(* IEC 61131-3 sources: stdmachine/plc/src/05_Sequencers (part 2) *)

(* ---- FB_Machine.st ---- *)
// Bloc de tête du PLC (docs/05 § 5.1, § 5.2, § 10 ; docs/06 § 6) : machine d'états de la machine, propagation des
// commandes aux stations, défauts machine et raison d'arrêt, objets de niveau machine, système planaire, séquenceur
// général, calibrations machine, chargeur, handshakes de GVL_Hmi, forçages, surveillance des rebuts, balise,
// identité du PLC, battement de la HMI, publication du statut.
//
// Le projet de la machine l'appelle une fois par cycle dans MAIN : fbMachine(); après avoir renseigné GVL_IoRef.
// Avant le premier appel, il peut donner ses pools (SetPools) et son pilote planaire (SetPlanarDriver) ; sinon la
// bibliothèque prend FB_DefaultPools et le système planaire simulé.
FUNCTION_BLOCK FB_Machine EXTENDS FB_NodeBase IMPLEMENTS I_ManualHost, I_ObjectHost
VAR
    fbPack : FB_PackML;
    aStation : ARRAY[1..GVL_Const.MAX_STATIONS] OF FB_Station;
    fbSeq : FB_GeneralSequencer;
    fbMgr : FB_MoverManager;
    fbPlanarSim : FB_PlanarSim;
    fbAlarms : FB_AlarmManager;
    fbTraces : FB_TraceBuffer;
    fbQuality : FB_QualityMonitor;
    fbFactory : FB_ObjectFactory;
    fbLoader : FB_Loader;
    fbCalib : FB_MachineCalib;
    fbDefaultPools : FB_DefaultPools;
    fbManual : FB_ManualChannel;            // canal 0 : objets de niveau machine
    _ipPools : I_ObjectPools;
    _ipPlanar : I_PlanarDriver;
    _bSimPlanar : BOOL;
    aObj : ARRAY[1..GVL_Const.MAX_MACHINE_OBJ] OF I_Object;
    _nObj : UINT;
    _bInit : BOOL;
    _ePendingCmd : E_Cmd;
    _sCmdUser : STRING(24);
    _eReasonNext : E_StopReason;            // cause système du prochain arrêt
    _bOperatorAwaited : BOOL;               // fin d'OF, machine vidée : bleu clignotant jusqu'au prochain Start
    // Handshakes (docs/06 § 6.1) : dernier nSeq traité
    _nCmdSeq : UDINT;
    _nOverrideSeq : UDINT;
    _nLaunchSeq : UDINT;
    _nOrderSeq : UDINT;
    _nMoverVarSeq : UDINT;
    _nPromptSeq : UDINT;
    _nPartSeq : UDINT;
    _nAckSeq : UDINT;
    _nForceSeq : UDINT;
    _nQualitySeq : UDINT;
    _nSimForceSeq : UDINT;
    // Battement de la HMI
    _nLastHmiBeat : UDINT;
    _fHmiQuietMs : LREAL;
    bHmiLost : BOOL;
    _nHeartbeat : UDINT;
    _fRetainedMs : LREAL;
    _tLastCalibCheck : LINT;
    _nPlanarError : UINT;
END_VAR
VAR PERSISTENT
    stForce : ST_MachineForce;              // forçages et état déclaré (docs/12)
    _fMachineOverride : LREAL := 100.0;
    _aStationOverride : ARRAY[1..GVL_Const.MAX_STATIONS] OF LREAL := [16(100.0)];
    _eMode : E_Mode;
    _nStopCauseGid : UDINT;
    _nStopCauseCode : UINT;
    _eStopReason : E_StopReason;
END_VAR

_Run();

// ================================================================== mise en place

METHOD SetPools
VAR_INPUT
    ipPools : I_ObjectPools;
END_VAR
_ipPools := ipPools;
END_METHOD

METHOD SetPlanarDriver
VAR_INPUT
    ipDriver : I_PlanarDriver;
END_VAR
_ipPlanar := ipDriver;
END_METHOD

METHOD PRIVATE _Init
VAR
    n : USINT;
    t : UINT;
    stResp : ST_DeployResponse;
END_VAR
fbAlarms.Bind(GVL_Hmi.stAlarms);
fbTraces.Bind(GVL_Hmi.stTraces);
IF _ipPools = 0 THEN _ipPools := fbDefaultPools; END_IF
IF _ipPlanar = 0 THEN
    _ipPlanar := fbPlanarSim;
    _bSimPlanar := TRUE;
END_IF
fbFactory.SetPools(_ipPools, fbAlarms);
fbFactory.SetHost(0, THIS^, THIS^, 0);
FOR n := 1 TO GVL_Const.MAX_STATIONS DO
    aStation[n].Init(nStation := n, refData := GVL_Active.aStation[n], refMachine := GVL_Active.stMachine, refAlarms := fbAlarms,
                     refStatus := GVL_Hmi.aStationStatus[n], refStep := GVL_Hmi.aStep[n], ipMachine := THIS^);
    aStation[n].SetOverride(_aStationOverride[n]);
    fbFactory.SetHost(n, aStation[n], aStation[n], aStation[n]);
    fbSeq.SetStation(n, ADR(aStation[n]));
    fbCalib.SetStation(n, ADR(aStation[n]));
END_FOR
fbQuality.Init(GVL_Active.stMachine, fbAlarms);
fbMgr.Init(GVL_Active.stMachine, _ipPlanar);
GVL_IoRef.ipPlanar := _ipPlanar;
GVL_IoRef.ipMovers := fbMgr;
fbSeq.Init(GVL_Active.stMachine, fbMgr, fbQuality, fbAlarms, fbTraces);
fbCalib.Init(GVL_Active.stMachine, fbAlarms, fbMgr);
fbManual.Init(nStation := 0, ipHost := THIS^);
fbLoader.Init(fbFactory);
SetOverride(_fMachineOverride);

// Mémoire rémanente : identifiant tiré à sa première initialisation (docs/02 § 7.4)
IF GVL_Active.nRetainId = 0 THEN
    GVL_Active.nRetainId := LINT_TO_ULINT(F_NowUtc()) XOR 16#9E3779B97F4A7C15;
END_IF

// Redémarrage du PLC : le dernier déploiement reste actif, les objets sont rattachés de nouveau à leurs éléments
IF GVL_Active.bDeployed THEN
    fbFactory.Build(stResp);
    fbMgr.Configure();
    fbSeq.ScanGroups();
    _PlaceSimMovers();
END_IF
FOR n := 1 TO GVL_Const.MAX_STATIONS DO aStation[n].SetMode(_eMode); END_FOR

// Identité (docs/05 § 10)
GVL_Hmi.stIdentity.nInterfaceVersion := GVL_Const.INTERFACE_VERSION;
GVL_Hmi.stIdentity.nInstrSetVersion := GVL_Const.INSTR_SET_VERSION;
GVL_Hmi.stIdentity.nCatalogVersion := GVL_Catalog.CatalogVersion;
GVL_Hmi.stIdentity.sLibVersion := GVL_Const.LIB_VERSION;
GVL_Hmi.stIdentity.nRetainId := GVL_Active.nRetainId;
FOR t := 1 TO GVL_Const.MAX_TYPE DO GVL_Hmi.stIdentity.aPoolSize[t] := fbFactory.PoolSize(t); END_FOR

// Les demandes déjà présentes dans GVL_Hmi au démarrage ne sont pas rejouées
_nCmdSeq := GVL_Hmi.stCmd.nSeq;
_nOverrideSeq := GVL_Hmi.stOverride.nSeq;
_nLaunchSeq := GVL_Hmi.stLaunch.nSeq;
_nOrderSeq := GVL_Hmi.stOrder.nSeq;
_nMoverVarSeq := GVL_Hmi.stMoverVar.nSeq;
_nPromptSeq := GVL_Hmi.stPrompt.nSeq;
_nPartSeq := GVL_Hmi.stPartCmd.nSeq;
_nAckSeq := GVL_Hmi.stAlarmAck.nSeq;
_nForceSeq := GVL_Hmi.stForceCmd.nSeq;
_nQualitySeq := GVL_Hmi.stQualityCmd.nSeq;
_nSimForceSeq := GVL_Hmi.stSimForce.nSeq;
_nLastHmiBeat := GVL_Hmi.nHmiHeartbeat;
_ApplyMoverForces();
_bInit := TRUE;
END_METHOD

// Simulation : chaque mover est posé sur une position tampon, sinon de parcage, sinon en ligne (docs/06 § 8)
METHOD PRIVATE _PlaceSimMovers
VAR
    i : USINT;
    k : INT;
    nPlaced : USINT;
    stPos : ST_Position;
END_VAR
IF NOT _bSimPlanar THEN RETURN; END_IF
fbPlanarSim.SetMoverCount(GVL_Active.stMachine.nMovers);
nPlaced := 0;
FOR k := 1 TO GVL_Active.stMachine.nPlanarPos DO
    IF nPlaced < GVL_Active.stMachine.nMovers AND (GVL_Active.stMachine.aPlanarPos[k].eKind = E_PlanarPosKind.Buffer
       OR GVL_Active.stMachine.aPlanarPos[k].eKind = E_PlanarPosKind.Park) THEN
        nPlaced := nPlaced + 1;
        fbPlanarSim.SetInitialPosition(nPlaced, GVL_Active.stMachine.aPlanarPos[k].stPos);
    END_IF
END_FOR
FOR i := nPlaced + 1 TO GVL_Active.stMachine.nMovers DO
    MEMSET(ADR(stPos), 0, SIZEOF(stPos));
    stPos.fX := USINT_TO_LREAL(i) * 120.0;
    fbPlanarSim.SetInitialPosition(i, stPos);
END_FOR
END_METHOD

// ================================================================== cycle

METHOD PRIVATE _Run
VAR
    n : USINT;
    k : UINT;
    eBefore : E_State;
    eCmd : E_Cmd;
    tNow : LINT;
END_VAR
IF NOT _bInit THEN _Init(); END_IF
tNow := F_NowUtc();
_nHeartbeat := _nHeartbeat + 1;
_WatchHmi();

// Chargeur : vérification, activation, restauration (machine Stopped)
fbLoader(bMachineStopped := fbPack.eState = E_State.Stopped);
fbLoader.Cycle();
IF fbLoader.bActivate THEN _Activate(); END_IF
IF fbLoader.bRestore THEN _ApplyRestore(); END_IF

// Demandes de la HMI
_HandleCmd();
_HandleOverride();
_HandleLaunch();
_HandleOrder();
_HandleMoverVar();
_HandlePrompt();
_HandlePart();
_HandleAlarmAck();
_HandleForce();
_HandleQuality();
_HandleSimForce();

// Arrêts automatiques demandés au cycle précédent : OF terminé, machine vidée, réaction qualité
IF fbSeq.bStopRequest AND _ePendingCmd = E_Cmd.None AND fbPack.Accepts(E_Cmd.Stop) THEN
    _ePendingCmd := E_Cmd.Stop;
    CASE fbSeq.nStopReason OF
        1: _eReasonNext := E_StopReason.OrderComplete;
        2: _eReasonNext := E_StopReason.Drained;
    ELSE
        _eReasonNext := E_StopReason.Quality;
    END_CASE
    _bOperatorAwaited := fbSeq.nStopReason <> 3;
END_IF

// Système planaire
UpdateOverride();
fbMgr.Cycle(EffectiveOverride);         // fait aussi tourner le pilote planaire
_PlanarAlarms();

// Machine d'états
eCmd := _ePendingCmd;
_ePendingCmd := E_Cmd.None;
eBefore := fbPack.eState;
fbPack(eCmd := eCmd, bStateComplete := _StateComplete(), bFault := _Fault());
IF fbPack.bEntry THEN _OnEntry(eBefore); END_IF

// Objets de niveau machine
_UpdateObjects();
fbManual.Cycle();

// Stations : forçages et réactions qualité, puis leur cycle
FOR n := 1 TO GVL_Const.MAX_STATIONS DO
    aStation[n].SetOutOfProduction(stForce.aStation[n].bOutOfProduction);
    aStation[n].SetQualityLock(fbQuality.aStationHold[n]);
    aStation[n].Cycle();
END_FOR

// Séquenceur général et calibration machine
fbSeq.Cycle(fbPack.eState);
IF fbCalib.bRunning AND (fbPack.eState <> E_State.Idle OR _eMode <> E_Mode.Maintenance) THEN fbCalib.Abort(); END_IF
fbCalib.Cycle(bHmiLost);

// Calibrations échues : une fois par jour (et à chaque Reset, voir _OnEntry)
IF tNow - _tLastCalibCheck > 864000000000 THEN _CheckCalibrations(tNow); END_IF

_Beacon();
fbQuality.Publish();
_fRetainedMs := _fRetainedMs + F_CycleMs();
IF _fRetainedMs >= 1000.0 THEN
    _fRetainedMs := 0;
    _PublishRetained();
END_IF
_Publish();
END_METHOD

METHOD PRIVATE _WatchHmi
IF GVL_Hmi.nHmiHeartbeat <> _nLastHmiBeat THEN
    _nLastHmiBeat := GVL_Hmi.nHmiHeartbeat;
    _fHmiQuietMs := 0;
    bHmiLost := FALSE;
ELSE
    _fHmiQuietMs := _fHmiQuietMs + F_CycleMs();
    IF _fHmiQuietMs >= GVL_Const.HMI_HEARTBEAT_MS AND NOT bHmiLost THEN
        bHmiLost := TRUE;
        fbAlarms.RaiseEvent(0, 917, 0, E_Severity.Info);           // la production continue (docs/06 § 6.2)
    END_IF
END_IF
END_METHOD

// ================================================================== machine d'états (docs/05 § 5.1 et 5.2)

METHOD PRIVATE _StateComplete : BOOL
VAR
    n : USINT;
    bAll : BOOL := TRUE;
END_VAR
_StateComplete := FALSE;
CASE fbPack.eState OF
    E_State.Resetting:
        // Système planaire actif, movers détectés (un mover hors service peut être absent), chaque fonction
        // utilisée a une station en Idle
        IF NOT _ipPlanar.Activate(TRUE) THEN RETURN; END_IF
        _StateComplete := _AllMoversDetected() AND fbSeq.MissingGroup(2) = 0;
    E_State.Stopping:
        FOR n := 1 TO GVL_Const.MAX_STATIONS DO
            IF aStation[n].State <> E_State.Stopped AND aStation[n].State <> E_State.Aborted THEN bAll := FALSE; END_IF
        END_FOR
        _StateComplete := bAll AND NOT fbMgr.AnyMoving();
    E_State.Clearing:
        FOR n := 1 TO GVL_Const.MAX_STATIONS DO
            IF aStation[n].State = E_State.Clearing THEN bAll := FALSE; END_IF
        END_FOR
        _StateComplete := bAll AND _ObjectsOk();
END_CASE
END_METHOD

METHOD PRIVATE _AllMoversDetected : BOOL
VAR
    i : USINT;
END_VAR
_AllMoversDetected := TRUE;
FOR i := 1 TO GVL_Active.stMachine.nMovers DO
    IF NOT _ipPlanar.MoverDetected(i) THEN
        IF NOT stForce.aMover[i].bOutOfService THEN
            _AllMoversDetected := FALSE;
            fbAlarms.Raise(_PlanarGlobalId(), 101, i, E_Severity.Warning);    // « Mover non détecté » : reste en Resetting
        END_IF
    ELSE
        fbAlarms.Clear(_PlanarGlobalId(), 101);
    END_IF
END_FOR
END_METHOD

METHOD PRIVATE _Fault : BOOL
VAR
    n : USINT;
    g : USINT;
    eSt : E_State;
    ipSafety : I_SafetyCircuits;
    k : UINT;
END_VAR
_Fault := FALSE;
eSt := fbPack.eState;
// Circuits de sécurité de niveau machine
FOR k := 1 TO _nObj DO
    IF aObj[k] <> 0 AND_THEN __QUERYINTERFACE(aObj[k], ipSafety) THEN
        IF NOT ipSafety.AllOk THEN _Fault := TRUE; END_IF
    END_IF
END_FOR
IF eSt = E_State.Stopped THEN RETURN; END_IF          // à l'arrêt, une sécurité ouverte n'est pas un défaut
// Système planaire, movers, alarmes de process de gravité défaut machine
IF _nPlanarError <> 0 OR fbSeq.bMachineFault THEN _Fault := TRUE; END_IF
IF eSt <> E_State.Aborted AND eSt <> E_State.Clearing THEN
    FOR n := 1 TO GVL_Const.MAX_STATIONS DO
        IF aStation[n].MachineFault THEN _Fault := TRUE; END_IF
    END_FOR
    IF NOT _ObjectsOk() THEN _Fault := TRUE; END_IF
END_IF
// Fonction utilisée sans station disponible (913) ; au Reset, fonction dont toutes les stations ont échoué
IF eSt = E_State.Execute THEN
    g := fbSeq.MissingGroup(1);
ELSIF eSt = E_State.Resetting THEN
    g := fbSeq.MissingGroup(3);
END_IF
IF g <> 0 THEN
    fbAlarms.RaiseEvent(0, 913, g, E_Severity.MachineFault);
    _Fault := TRUE;
END_IF
END_METHOD

METHOD PRIVATE _ObjectsOk : BOOL
VAR
    k : UINT;
END_VAR
_ObjectsOk := TRUE;
FOR k := 1 TO _nObj DO
    IF aObj[k] <> 0 THEN
        IF aObj[k].NodeState = E_ObjState.Error THEN _ObjectsOk := FALSE; END_IF
    END_IF
END_FOR
END_METHOD

METHOD PRIVATE _OnEntry
VAR_INPUT
    eFrom : E_State;
END_VAR
VAR
    n : USINT;
    k : UINT;
    eSt : E_State;
END_VAR
CASE fbPack.eState OF
    E_State.Stopped:
        fbSeq.bDrain := FALSE;
    E_State.Resetting:
        _ClearStopCause();
        FOR k := 1 TO _nObj DO IF aObj[k] <> 0 THEN aObj[k].Ack(); END_IF END_FOR
        _ipPlanar.AckError();
        FOR n := 1 TO GVL_Const.MAX_STATIONS DO
            IF _StationUsed(n) AND aStation[n].State = E_State.Stopped THEN aStation[n].Command(E_Cmd.Reset); END_IF
        END_FOR
        _CheckCalibrations(F_NowUtc());
    E_State.Idle:
        // Fin du Reset : chaque mover reçoit sa position, contextes et pièces gardés (docs/05 § 6.3)
        IF eFrom = E_State.Resetting THEN fbSeq.OnReset(); END_IF
    E_State.Execute:
        _ClearStopCause();
        _bOperatorAwaited := FALSE;
        FOR n := 1 TO GVL_Const.MAX_STATIONS DO
            eSt := aStation[n].State;
            IF _StationUsed(n) AND (eSt = E_State.Idle OR eSt = E_State.Held) THEN aStation[n].Command(E_Cmd.Start); END_IF
        END_FOR
    E_State.Held:
        _TakeStopCause();
        FOR n := 1 TO GVL_Const.MAX_STATIONS DO
            IF aStation[n].State = E_State.Execute THEN aStation[n].Command(E_Cmd.Hold); END_IF
        END_FOR
    E_State.Stopping:
        _TakeStopCause();
        fbSeq.bDrain := FALSE;
        FOR n := 1 TO GVL_Const.MAX_STATIONS DO
            eSt := aStation[n].State;
            IF eSt = E_State.Resetting OR eSt = E_State.Idle OR eSt = E_State.Execute OR eSt = E_State.Held THEN aStation[n].Command(E_Cmd.Stop); END_IF
        END_FOR
    E_State.Aborted:
        _TakeStopCause();
        fbSeq.bDrain := FALSE;
        fbMgr.StopAll();
        fbCalib.Abort();
        FOR k := _nObj TO 1 BY -1 DO IF aObj[k] <> 0 THEN aObj[k].Abort(); END_IF END_FOR
        FOR n := 1 TO GVL_Const.MAX_STATIONS DO
            IF aStation[n].State <> E_State.Aborted AND aStation[n].State <> E_State.Stopped THEN aStation[n].Command(E_Cmd.Abort); END_IF
        END_FOR
    E_State.Clearing:
        fbAlarms.AckFaults(0, FALSE, _sCmdUser);
        FOR k := 1 TO _nObj DO IF aObj[k] <> 0 THEN aObj[k].Ack(); END_IF END_FOR
        fbSeq.ClearFaults();
        _ipPlanar.AckError();
        FOR n := 1 TO GVL_Const.MAX_STATIONS DO
            IF aStation[n].State = E_State.Aborted THEN aStation[n].Command(E_Cmd.Clear); END_IF
        END_FOR
END_CASE
END_METHOD

METHOD PRIVATE _StationUsed : BOOL
VAR_INPUT
    n : USINT;
END_VAR
_StationUsed := GVL_Active.stMachine.aStation[n].bUsed;
END_METHOD

// Raison d'arrêt (docs/05 § 5.2, docs/14 § 4) : première alarme cause, sinon la cause système
METHOD PRIVATE _TakeStopCause
VAR
    i : INT;
END_VAR
IF _eStopReason <> E_StopReason.None THEN RETURN; END_IF      // déjà prise pour cet épisode d'arrêt
// Un arrêt automatique (OF terminé, machine vidée, qualité) garde sa cause même si une alarme est active
IF _eReasonNext = E_StopReason.OrderComplete OR _eReasonNext = E_StopReason.Drained OR _eReasonNext = E_StopReason.Quality THEN
    _eStopReason := _eReasonNext;
    _eReasonNext := E_StopReason.None;
    RETURN;
END_IF
i := fbAlarms.FirstFault(0, TRUE);
IF i > 0 THEN
    fbAlarms.MarkCause(i);
    _nStopCauseGid := GVL_Hmi.stAlarms.aActive[i].nGlobalId;
    _nStopCauseCode := GVL_Hmi.stAlarms.aActive[i].nCode;
    _eStopReason := E_StopReason.Alarm;
ELSE
    _eStopReason := E_StopReason.Operator;
END_IF
_eReasonNext := E_StopReason.None;
END_METHOD

METHOD PRIVATE _ClearStopCause
_nStopCauseGid := 0;
_nStopCauseCode := 0;
_eStopReason := E_StopReason.None;
_eReasonNext := E_StopReason.None;
END_METHOD

METHOD PRIVATE _CheckCalibrations
VAR_INPUT
    tNow : LINT;
END_VAR
VAR
    n : USINT;
END_VAR
_tLastCalibCheck := tNow;
FOR n := 1 TO GVL_Const.MAX_STATIONS DO
    IF _StationUsed(n) THEN aStation[n].CheckCalibrations(tNow); END_IF
END_FOR
fbCalib.CheckCalibrations(tNow);
END_METHOD

// ================================================================== système planaire et objets machine

METHOD PRIVATE _PlanarGlobalId : UDINT
VAR
    k : UINT;
END_VAR
_PlanarGlobalId := 0;
FOR k := 1 TO MIN(GVL_Active.stMachine.nMachineObj, GVL_Const.MAX_MACHINE_OBJ) DO
    IF GVL_Active.stMachine.aMachineObj[k].nType = GVL_Catalog.Type_PlanarSystem THEN
        _PlanarGlobalId := UINT_TO_UDINT(GVL_Active.stMachine.aMachineObj[k].nLocalId);
        RETURN;
    END_IF
END_FOR
END_METHOD

METHOD PRIVATE _PlanarAlarms
VAR
    nErr : UINT;
END_VAR
nErr := _ipPlanar.ErrorCode;
IF nErr <> _nPlanarError THEN
    IF _nPlanarError <> 0 THEN fbAlarms.Clear(_PlanarGlobalId(), _nPlanarError); END_IF
    IF nErr <> 0 THEN fbAlarms.Raise(_PlanarGlobalId(), nErr, _ipPlanar.ErrorSubCode, E_Severity.MachineFault); END_IF
    _nPlanarError := nErr;
END_IF
END_METHOD

METHOD PRIVATE _UpdateObjects
VAR
    k : UINT;
END_VAR
FOR k := 1 TO _nObj DO
    IF aObj[k] <> 0 THEN
        aObj[k].Cycle();
        GVL_Hmi.aObjStatus[0, k] := aObj[k].Status;
    END_IF
END_FOR
END_METHOD

// Balise de la machine (docs/02 § 8) : pilotée par l'état de la machine
METHOD PRIVATE _Beacon
VAR
    k : UINT;
    n : USINT;
    nPattern : UINT;
    bMaint : BOOL;
    bStationAborted : BOOL;
    ipBeacon : I_Beacon;
END_VAR
bMaint := _eMode = E_Mode.Maintenance OR stForce.eDeclared = E_DeclaredState.PlannedMaintenance
          OR stForce.eDeclared = E_DeclaredState.CorrectiveMaintenance OR stForce.eDeclared = E_DeclaredState.Trials
          OR stForce.eDeclared = E_DeclaredState.Cleaning;
FOR n := 1 TO GVL_Const.MAX_STATIONS DO
    IF aStation[n].State = E_State.Aborted THEN bStationAborted := TRUE; END_IF
END_FOR
nPattern := F_BeaconPattern(fbPack.eState, bMaint, _bOperatorAwaited OR fbSeq.AnyToEmpty() OR fbQuality.bAnyReaction, bStationAborted);
FOR k := 1 TO _nObj DO
    IF aObj[k] <> 0 AND_THEN __QUERYINTERFACE(aObj[k], ipBeacon) THEN ipBeacon.SetPattern(nPattern, (nPattern AND GVL_BeaconBits.BUZZER) <> 0); END_IF
END_FOR
END_METHOD

// ================================================================== déploiement (docs/05 § 10)

METHOD PRIVATE _Activate
VAR
    stResp : ST_DeployResponse;
    n : USINT;
    nOldGeneral : INT;
    nNewGeneral : INT;
    bRestart : BOOL;
END_VAR
IF fbPack.eState <> E_State.Stopped THEN
    F_AddDeployError(stResp, 21, 0, 0, 0, 0, 0);
    fbLoader.Finish(stResp);
    RETURN;
END_IF
nOldGeneral := _GeneralSize(GVL_Active.stMachine);
nNewGeneral := _GeneralSize(GVL_Hmi.stStaging.stMachine);
bRestart := NOT GVL_Active.bDeployed OR nOldGeneral <> nNewGeneral
            OR GVL_Active.stMachine.nMovers <> GVL_Hmi.stStaging.stMachine.nMovers
            OR GVL_Active.stMachine.nSlots <> GVL_Hmi.stStaging.stMachine.nSlots;
// Copie atomique de la zone d'attente (un seul cycle)
GVL_Active.stMachine := GVL_Hmi.stStaging.stMachine;
GVL_Active.aStation := GVL_Hmi.stStaging.aStation;
GVL_Active.aPressRecipe := GVL_Hmi.stStaging.aPressRecipe;
GVL_Active.stMachine.tDeployed := F_NowUtc();
GVL_Active.stMachine.sDeployedBy := fbLoader.Request.sUser;
GVL_Active.bDeployed := TRUE;
fbFactory.Build(stResp);
FOR n := 1 TO GVL_Const.MAX_STATIONS DO aStation[n].OnDeploy(); END_FOR
fbMgr.Configure();
fbSeq.OnDeploy(bRestart);
fbCalib.OnDeploy();
_PlaceSimMovers();
fbLoader.Finish(stResp);
END_METHOD

// Taille du process général : somme des longueurs de ses tables (docs/05 § 10, étape 4)
METHOD PRIVATE _GeneralSize : INT
VAR_IN_OUT
    stData : ST_MachineData;
END_VAR
VAR
    t : USINT;
END_VAR
_GeneralSize := 0;
FOR t := 1 TO GVL_Const.MAX_TABLES DO
    IF stData.aTable[t].bUsed AND (stData.aTable[t].eKind = E_TableKind.General OR stData.aTable[t].eKind = E_TableKind.GeneralSub) THEN
        _GeneralSize := _GeneralSize + stData.aTable[t].nLength;
    END_IF
END_FOR
END_METHOD

// Restauration des valeurs rémanentes (docs/05 § 10, étape 6)
METHOD PRIVATE _ApplyRestore
VAR
    k : UINT;
    nUnknown : UINT;
    stItem : ST_RetainedItem;
    bOk : BOOL;
END_VAR
FOR k := 1 TO fbLoader.nRestoreCount DO
    stItem := fbLoader.aRestore[k];
    bOk := FALSE;
    CASE stItem.eKind OF
        E_RetainedKind.StationVar:
            IF stItem.nStation >= 1 AND stItem.nStation <= GVL_Const.MAX_STATIONS THEN bOk := aStation[stItem.nStation].Restore(stItem); END_IF
        E_RetainedKind.Calibration:
            IF stItem.nStation = 0 THEN
                bOk := fbCalib.Restore(stItem);
            ELSIF stItem.nStation <= GVL_Const.MAX_STATIONS THEN
                bOk := aStation[stItem.nStation].Restore(stItem);
            END_IF
        E_RetainedKind.MoverVar:
            bOk := fbSeq.Restore(stItem);
        E_RetainedKind.ObjectCounters:
            bOk := fbFactory.Restore(stItem);
    END_CASE
    IF NOT bOk THEN nUnknown := nUnknown + 1; END_IF          // compteurs de production : avec FB_PlantPublisher
END_FOR
fbLoader.RestoreDone(nUnknown);
_PublishRetained();
END_METHOD

METHOD PRIVATE _PublishRetained
VAR
    n : USINT;
END_VAR
GVL_Hmi.stRetained.nRetainId := GVL_Active.nRetainId;
GVL_Hmi.stRetained.nCount := 0;
FOR n := 1 TO GVL_Const.MAX_STATIONS DO
    IF _StationUsed(n) THEN aStation[n].PublishRetained(GVL_Hmi.stRetained); END_IF
END_FOR
fbCalib.PublishRetained(GVL_Hmi.stRetained);
fbSeq.PublishRetained(GVL_Hmi.stRetained);
fbFactory.PublishRetained(GVL_Hmi.stRetained);
END_METHOD

// ================================================================== demandes de la HMI (docs/06 § 6.2)

METHOD PRIVATE _HandleCmd
VAR
    req : REFERENCE TO ST_CmdRequest;
    resp : REFERENCE TO ST_CmdResponse;
    n : USINT;
    eReason : E_RejectReason;
    eSt : E_State;
END_VAR
req REF= GVL_Hmi.stCmd;
resp REF= GVL_Hmi.stCmdResp;
IF req.nSeq = _nCmdSeq THEN RETURN; END_IF
_nCmdSeq := req.nSeq;
eReason := E_RejectReason.None;
IF req.nTarget = 0 THEN
    IF req.bSetMode THEN
        eReason := _SetMode(req.eMode);
    ELSE
        eReason := _MachineCommand(req.eCmd, req.sUser);
    END_IF
    resp.eState := fbPack.eState;
ELSIF req.nTarget > GVL_Const.MAX_STATIONS OR_ELSE NOT _StationUsed(req.nTarget) THEN
    eReason := E_RejectReason.NotConfigured;
ELSE
    // Commande d'une station seule : réintégration pendant que la machine produit (docs/05 § 5.1)
    n := req.nTarget;
    eSt := aStation[n].State;
    IF req.bSetMode THEN
        eReason := E_RejectReason.NotAllowed;       // le mode est celui de la machine
    ELSIF NOT (fbPack.eState = E_State.Execute OR fbPack.eState = E_State.Held) THEN
        eReason := E_RejectReason.WrongState;
    ELSIF (eSt = E_State.Execute OR eSt = E_State.Held) AND NOT aStation[n].OutOfProduction THEN
        eReason := E_RejectReason.NotAllowed;       // station en production : elle suit la machine
    ELSE
        eReason := aStation[n].Command(req.eCmd);
    END_IF
    resp.eState := eSt;
END_IF
resp.eReason := eReason;
resp.eResult := SEL(eReason = E_RejectReason.None, E_CmdResult.Rejected, E_CmdResult.Accepted);
resp.nDetail := 0;
resp.nSeq := req.nSeq;
END_METHOD

METHOD PRIVATE _MachineCommand : E_RejectReason
VAR_INPUT
    eCmd : E_Cmd;
    sUser : STRING(24);
END_VAR
VAR
    eSt : E_State;
END_VAR
eSt := fbPack.eState;
_MachineCommand := E_RejectReason.None;
CASE eCmd OF
    E_Cmd.DrainStart:
        IF eSt = E_State.Execute OR eSt = E_State.Held OR eSt = E_State.Idle THEN fbSeq.bDrain := TRUE;
        ELSE _MachineCommand := E_RejectReason.WrongState; END_IF
        RETURN;
    E_Cmd.DrainCancel:
        fbSeq.bDrain := FALSE;
        RETURN;
    E_Cmd.Start:
        IF stForce.bStartBlocked THEN _MachineCommand := E_RejectReason.StartBlocked; RETURN; END_IF
    E_Cmd.Reset:
        IF NOT GVL_Active.bDeployed THEN _MachineCommand := E_RejectReason.NotConfigured; RETURN; END_IF
        IF fbLoader.bBusy THEN _MachineCommand := E_RejectReason.Busy; RETURN; END_IF
END_CASE
IF eCmd = E_Cmd.None OR NOT fbPack.Accepts(eCmd) THEN
    _MachineCommand := E_RejectReason.WrongState;
    RETURN;
END_IF
_ePendingCmd := eCmd;
_sCmdUser := sUser;
IF eCmd = E_Cmd.Stop OR eCmd = E_Cmd.Hold OR eCmd = E_Cmd.Abort THEN _eReasonNext := E_StopReason.Operator; END_IF
END_METHOD

METHOD PRIVATE _SetMode : E_RejectReason
VAR_INPUT
    eMode : E_Mode;
END_VAR
VAR
    n : USINT;
END_VAR
IF fbPack.eState <> E_State.Stopped THEN _SetMode := E_RejectReason.WrongState; RETURN; END_IF
FOR n := 1 TO GVL_Const.MAX_STATIONS DO
    IF aStation[n].State <> E_State.Stopped THEN _SetMode := E_RejectReason.WrongState; RETURN; END_IF
END_FOR
_eMode := eMode;
FOR n := 1 TO GVL_Const.MAX_STATIONS DO aStation[n].SetMode(eMode); END_FOR
_SetMode := E_RejectReason.None;
END_METHOD

METHOD PRIVATE _HandleOverride
VAR
    req : REFERENCE TO ST_OverrideRequest;
    resp : REFERENCE TO ST_CmdResponse;
END_VAR
req REF= GVL_Hmi.stOverride;
resp REF= GVL_Hmi.stOverrideResp;
IF req.nSeq = _nOverrideSeq THEN RETURN; END_IF
_nOverrideSeq := req.nSeq;
resp.eReason := E_RejectReason.None;
IF req.nObject <> 0 OR req.bManual THEN
    resp.eReason := E_RejectReason.NotAllowed;          // override d'objet : propriété de la configuration (D94)
ELSIF req.nStation = 0 THEN
    _fMachineOverride := LIMIT(0.0, req.fValue, 100.0);
    SetOverride(_fMachineOverride);
ELSIF req.nStation <= GVL_Const.MAX_STATIONS THEN
    _aStationOverride[req.nStation] := LIMIT(0.0, req.fValue, 100.0);
    aStation[req.nStation].SetOverride(_aStationOverride[req.nStation]);
ELSE
    resp.eReason := E_RejectReason.NotConfigured;
END_IF
resp.eResult := SEL(resp.eReason = E_RejectReason.None, E_CmdResult.Rejected, E_CmdResult.Accepted);
resp.eState := fbPack.eState;
resp.nSeq := req.nSeq;
END_METHOD

METHOD PRIVATE _HandleLaunch
VAR
    req : REFERENCE TO ST_LaunchRequest;
    resp : REFERENCE TO ST_CmdResponse;
    pMover : POINTER TO ST_MoverCtx;
END_VAR
req REF= GVL_Hmi.stLaunch;
resp REF= GVL_Hmi.stLaunchResp;
IF req.nSeq = _nLaunchSeq THEN RETURN; END_IF
_nLaunchSeq := req.nSeq;
pMover := fbSeq.MoverPtr(req.nMover);
IF _eMode <> E_Mode.Maintenance THEN
    resp.eReason := E_RejectReason.WrongMode;
ELSIF req.nStation = 0 THEN
    // Calibration machine : machine Idle (docs/05 § 10.1)
    IF fbPack.eState <> E_State.Idle THEN resp.eReason := E_RejectReason.WrongState;
    ELSE resp.eReason := fbCalib.Start(req.nTable, req.nMover, pMover, req.sUser); END_IF
ELSIF req.nStation > GVL_Const.MAX_STATIONS OR_ELSE NOT _StationUsed(req.nStation) THEN
    resp.eReason := E_RejectReason.NotConfigured;
ELSE
    resp.eReason := aStation[req.nStation].Launch(req.nTable, req.nMover, pMover, req.nSlot, req.aParam, req.sUser);
END_IF
resp.eResult := SEL(resp.eReason = E_RejectReason.None, E_CmdResult.Rejected, E_CmdResult.Accepted);
resp.eState := fbPack.eState;
resp.nSeq := req.nSeq;
END_METHOD

METHOD PRIVATE _HandleOrder
VAR
    req : REFERENCE TO ST_OrderRequest;
    resp : REFERENCE TO ST_CmdResponse;
    eSt : E_State;
END_VAR
req REF= GVL_Hmi.stOrder;
resp REF= GVL_Hmi.stOrderResp;
IF req.nSeq = _nOrderSeq THEN RETURN; END_IF
_nOrderSeq := req.nSeq;
eSt := fbPack.eState;
CASE req.eCmd OF
    E_OrderCmd.Activate:
        IF eSt = E_State.Aborted OR eSt = E_State.Clearing OR eSt = E_State.Resetting OR eSt = E_State.Stopping THEN
            resp.eReason := E_RejectReason.WrongState;
        ELSE
            resp.eReason := fbSeq.Activate(req);
        END_IF
    E_OrderCmd.Suspend:
        resp.eReason := fbSeq.Suspend();
    E_OrderCmd.Cancel:
        resp.eReason := fbSeq.Cancel(req.nOrder);
ELSE
    resp.eReason := E_RejectReason.NotAllowed;
END_CASE
resp.eResult := SEL(resp.eReason = E_RejectReason.None, E_CmdResult.Rejected, E_CmdResult.Accepted);
resp.eState := eSt;
resp.nDetail := req.nOrder;
resp.nSeq := req.nSeq;
END_METHOD

METHOD PRIVATE _HandleMoverVar
VAR
    req : REFERENCE TO ST_MoverVarRequest;
    resp : REFERENCE TO ST_CmdResponse;
END_VAR
req REF= GVL_Hmi.stMoverVar;
resp REF= GVL_Hmi.stMoverVarResp;
IF req.nSeq = _nMoverVarSeq THEN RETURN; END_IF
_nMoverVarSeq := req.nSeq;
IF _eMode <> E_Mode.Maintenance THEN
    resp.eReason := E_RejectReason.WrongMode;
ELSIF fbPack.eState <> E_State.Stopped AND fbPack.eState <> E_State.Idle THEN
    resp.eReason := E_RejectReason.WrongState;
ELSE
    resp.eReason := fbSeq.SetMoverVar(req);
END_IF
resp.eResult := SEL(resp.eReason = E_RejectReason.None, E_CmdResult.Rejected, E_CmdResult.Accepted);
resp.eState := fbPack.eState;
resp.nSeq := req.nSeq;
END_METHOD

METHOD PRIVATE _HandlePrompt
VAR
    req : REFERENCE TO ST_PromptAnswer;
    resp : REFERENCE TO ST_CmdResponse;
    bOk : BOOL;
END_VAR
req REF= GVL_Hmi.stPrompt;
resp REF= GVL_Hmi.stPromptResp;
IF req.nSeq = _nPromptSeq THEN RETURN; END_IF
_nPromptSeq := req.nSeq;
IF req.nStation = 0 THEN
    bOk := fbCalib.AnswerPrompt(req.nPromptId, req.bConfirm);
ELSIF req.nStation <= GVL_Const.MAX_STATIONS THEN
    bOk := aStation[req.nStation].AnswerPrompt(req.nPromptId, req.bConfirm, req.fValue);
END_IF
resp.eReason := SEL(bOk, E_RejectReason.NotAllowed, E_RejectReason.None);
resp.eResult := SEL(bOk, E_CmdResult.Rejected, E_CmdResult.Accepted);
resp.eState := fbPack.eState;
resp.nSeq := req.nSeq;
END_METHOD

METHOD PRIVATE _HandlePart
VAR
    req : REFERENCE TO ST_PartRequest;
    resp : REFERENCE TO ST_CmdResponse;
END_VAR
req REF= GVL_Hmi.stPartCmd;
resp REF= GVL_Hmi.stPartResp;
IF req.nSeq = _nPartSeq THEN RETURN; END_IF
_nPartSeq := req.nSeq;
resp.eReason := fbSeq.ConfirmRemoved(req.nMover);
resp.eResult := SEL(resp.eReason = E_RejectReason.None, E_CmdResult.Rejected, E_CmdResult.Accepted);
resp.eState := fbPack.eState;
resp.nDetail := req.nMover;
resp.nSeq := req.nSeq;
END_METHOD

// Acquittement par l'opérateur : avertissements seulement ; les défauts s'acquittent par Clear (docs/14 § 4)
METHOD PRIVATE _HandleAlarmAck
VAR
    req : REFERENCE TO ST_AlarmAckRequest;
    resp : REFERENCE TO ST_CmdResponse;
END_VAR
req REF= GVL_Hmi.stAlarmAck;
resp REF= GVL_Hmi.stAlarmAckResp;
IF req.nSeq = _nAckSeq THEN RETURN; END_IF
_nAckSeq := req.nSeq;
fbAlarms.AckWarning(req.nGlobalId, req.nCode, req.sUser);
resp.eReason := E_RejectReason.None;
resp.eResult := E_CmdResult.Accepted;
resp.eState := fbPack.eState;
resp.nSeq := req.nSeq;
END_METHOD

// Forçages et état déclaré (docs/12) : mémorisés en persistant, publiés dans GVL_Hmi.stForce
METHOD PRIVATE _HandleForce
VAR
    req : REFERENCE TO ST_ForceCommand;
    resp : REFERENCE TO ST_CmdResponse;
    n : USINT;
END_VAR
req REF= GVL_Hmi.stForceCmd;
resp REF= GVL_Hmi.stForceResp;
IF req.nSeq = _nForceSeq THEN RETURN; END_IF
_nForceSeq := req.nSeq;
resp.eReason := E_RejectReason.None;
n := req.nTarget;
CASE req.eKind OF
    E_ForceKind.DeclaredState:
        IF req.bSet THEN
            stForce.eDeclared := req.eDeclared;
            stForce.bStartBlocked := req.bStartBlocked;
            stForce.nReason := req.nReason;
            stForce.tSince := F_NowUtc();
            stForce.tUntil := req.tUntil;
            stForce.sBy := req.sUser;
        ELSE
            stForce.eDeclared := E_DeclaredState.None;
            stForce.bStartBlocked := FALSE;
            stForce.nReason := 0;
            stForce.tSince := F_NowUtc();
            stForce.tUntil := 0;
            stForce.sBy := req.sUser;
        END_IF
    E_ForceKind.StationOutOfProduction:
        IF n < 1 OR n > GVL_Const.MAX_STATIONS OR_ELSE NOT _StationUsed(n) THEN
            resp.eReason := E_RejectReason.NotConfigured;
        ELSE
            stForce.aStation[n].bOutOfProduction := req.bSet;
            stForce.aStation[n].nReason := SEL(req.bSet, 0, req.nReason);
            stForce.aStation[n].tSince := F_NowUtc();
            stForce.aStation[n].sBy := req.sUser;
        END_IF
    E_ForceKind.MoverOutOfService:
        IF n < 1 OR n > GVL_Active.stMachine.nMovers THEN
            resp.eReason := E_RejectReason.NotConfigured;
        ELSE
            stForce.aMover[n].bOutOfService := req.bSet;
            stForce.aMover[n].bImmediate := req.bSet AND req.bImmediate;
            stForce.aMover[n].nReason := SEL(req.bSet, 0, req.nReason);
            stForce.aMover[n].tSince := F_NowUtc();
            stForce.aMover[n].sBy := req.sUser;
            fbSeq.SetOutOfService(n, req.bSet, req.bImmediate);
        END_IF
ELSE
    resp.eReason := E_RejectReason.NotAllowed;
END_CASE
resp.eResult := SEL(resp.eReason = E_RejectReason.None, E_CmdResult.Rejected, E_CmdResult.Accepted);
resp.eState := fbPack.eState;
resp.nSeq := req.nSeq;
END_METHOD

METHOD PRIVATE _ApplyMoverForces
VAR
    i : USINT;
END_VAR
FOR i := 1 TO GVL_Const.MAX_MOVERS DO
    fbSeq.SetOutOfService(i, stForce.aMover[i].bOutOfService, stForce.aMover[i].bImmediate);
END_FOR
END_METHOD

METHOD PRIVATE _HandleQuality
VAR
    req : REFERENCE TO ST_QualityCommand;
    resp : REFERENCE TO ST_CmdResponse;
END_VAR
req REF= GVL_Hmi.stQualityCmd;
resp REF= GVL_Hmi.stQualityResp;
IF req.nSeq = _nQualitySeq THEN RETURN; END_IF
_nQualitySeq := req.nSeq;
resp.eReason := E_RejectReason.None;
CASE req.eCmd OF
    E_QualityCmd.Release:
        IF NOT fbQuality.Release(req.eScope, req.nIndex) THEN resp.eReason := E_RejectReason.WrongState; END_IF
    E_QualityCmd.Reset:
        fbQuality.Reset(req.eScope, req.nIndex);
ELSE
    resp.eReason := E_RejectReason.NotAllowed;
END_CASE
resp.eResult := SEL(resp.eReason = E_RejectReason.None, E_CmdResult.Rejected, E_CmdResult.Accepted);
resp.eState := fbPack.eState;
resp.nSeq := req.nSeq;
END_METHOD

// Simulation : forcer une entrée simulée d'un objet (docs/12 § 5)
METHOD PRIVATE _HandleSimForce
VAR
    req : REFERENCE TO ST_SimForceRequest;
    resp : REFERENCE TO ST_CmdResponse;
    ipObj : I_Object;
END_VAR
req REF= GVL_Hmi.stSimForce;
resp REF= GVL_Hmi.stSimForceResp;
IF req.nSeq = _nSimForceSeq THEN RETURN; END_IF
_nSimForceSeq := req.nSeq;
IF req.nStation = 0 THEN
    ipObj := ObjectAt(req.nObject);
ELSIF req.nStation <= GVL_Const.MAX_STATIONS THEN
    ipObj := aStation[req.nStation].ObjectAt(req.nObject);
END_IF
IF ipObj = 0 THEN
    resp.eReason := E_RejectReason.NotConfigured;
ELSIF req.bRelease THEN
    ipObj.ForceInput(0, 0);
    resp.eReason := E_RejectReason.None;
ELSE
    ipObj.ForceInput(req.nSignal, req.fValue);
    resp.eReason := E_RejectReason.None;
END_IF
resp.eResult := SEL(resp.eReason = E_RejectReason.None, E_CmdResult.Rejected, E_CmdResult.Accepted);
resp.eState := fbPack.eState;
resp.nSeq := req.nSeq;
END_METHOD

// ================================================================== publication (docs/06 § 6.3)

METHOD PRIVATE _Publish
VAR
    s : REFERENCE TO ST_MachineStatus;
END_VAR
s REF= GVL_Hmi.stMachineStatus;
s.eState := fbPack.eState;
s.eMode := _eMode;
s.fEffOverride := LREAL_TO_REAL(EffectiveOverride);
s.nBeacon := F_BeaconPattern(fbPack.eState, _eMode = E_Mode.Maintenance, _bOperatorAwaited OR fbSeq.AnyToEmpty() OR fbQuality.bAnyReaction, FALSE);
s.bFault := fbPack.eState = E_State.Aborted;
s.tStateSince := fbPack.tSince;
s.nStopCauseGlobalId := _nStopCauseGid;
s.nStopCauseCode := _nStopCauseCode;
s.eStopReason := _eStopReason;
fbSeq.PublishOrders(s);
s.bDrain := fbSeq.bDrain;
s.nPartsInProcess := fbSeq.PartsInProcess();
s.bLoadingLocked := fbQuality.bLoadingLocked;
s.eDeclared := stForce.eDeclared;
s.bStartBlocked := stForce.bStartBlocked;
s.tPlcClock := F_NowUtc();
s.nPlcHeartbeat := _nHeartbeat;
s.sProjectHash := GVL_Active.stMachine.sProjectHash;
s.tDeployed := GVL_Active.stMachine.tDeployed;
s.bHmiLost := bHmiLost;
fbCalib.Publish(s);
GVL_Hmi.stForce := stForce;
END_METHOD

// ================================================================== I_ManualHost, I_ObjectHost

METHOD ObjectAt : I_Object
VAR_INPUT
    nLocalId : UINT;
END_VAR
IF nLocalId >= 1 AND nLocalId <= GVL_Const.MAX_MACHINE_OBJ THEN ObjectAt := aObj[nLocalId]; END_IF
END_METHOD

METHOD NamedPos : POINTER TO ST_NamedPos
VAR_INPUT
    nIndex : INT;
END_VAR
NamedPos := 0;                      // la machine n'a pas de positions nommées
END_METHOD

PROPERTY State : E_State
GET
State := fbPack.eState;
END_GET
END_PROPERTY

PROPERTY Mode : E_Mode
GET
Mode := _eMode;
END_GET
END_PROPERTY

METHOD ClearObjects
VAR
    k : UINT;
END_VAR
FOR k := 1 TO GVL_Const.MAX_MACHINE_OBJ DO aObj[k] := 0; END_FOR
_nObj := 0;
END_METHOD

METHOD SetObject
VAR_INPUT
    nLocalId : UINT;
    ipObj : I_Object;
END_VAR
IF nLocalId >= 1 AND nLocalId <= GVL_Const.MAX_MACHINE_OBJ THEN
    aObj[nLocalId] := ipObj;
    _nObj := MAX(_nObj, nLocalId);
END_IF
END_METHOD
END_FUNCTION_BLOCK

(* ---- FB_MachineCalib.st ---- *)
// Calibration machine (docs/05 § 10.1) : contexte unique, en Maintenance, machine Idle. Instructions reconnues :
// CalibStation (lance la calibration d'une station et l'attend), Route (le mover choisi au lancement seulement),
// Prompt, WaitTime, Jump, Alarm, End et les marqueurs ; toute autre instruction échoue (905).
FUNCTION_BLOCK FB_MachineCalib
VAR_OUTPUT
    bRunning : BOOL;
END_VAR
VAR
    _refMachine : REFERENCE TO ST_MachineData;
    _refAlarms : REFERENCE TO FB_AlarmManager;
    _refMgr : REFERENCE TO FB_MoverManager;
    aStation : ARRAY[1..GVL_Const.MAX_STATIONS] OF POINTER TO FB_Station;
    _nTable : INT;
    _nCalib : USINT;                // rang dans la liste des calibrations machine, 0 = table lancée sans déclaration
    _nPC : INT;
    _nWait : USINT;                 // 0 aucune, 1 durée, 2 station, 3 demande, 4 déplacement
    _fWaitMs : LREAL;
    _fElapsedMs : LREAL;
    _nStation : USINT;
    _nRetry : USINT;
    _nMover : USINT;
    _pMover : POINTER TO ST_MoverCtx;
    _nDest : INT;
    _sUser : STRING(24);
    stPrompt : ST_PromptState;
    _nPromptSeq : UDINT;
    _bAnswered : BOOL;
    _bConfirm : BOOL;
END_VAR
VAR PERSISTENT
    aCalib : ARRAY[1..GVL_Const.CALIB_PER_STATION] OF ST_CalibStatus;
END_VAR

METHOD Init
VAR_INPUT
    refMachine : REFERENCE TO ST_MachineData;
    refAlarms : REFERENCE TO FB_AlarmManager;
    refMgr : REFERENCE TO FB_MoverManager;
END_VAR
_refMachine REF= refMachine;
_refAlarms REF= refAlarms;
_refMgr REF= refMgr;
END_METHOD

METHOD SetStation
VAR_INPUT
    nStation : USINT;
    pStation : POINTER TO FB_Station;
END_VAR
IF nStation >= 1 AND nStation <= GVL_Const.MAX_STATIONS THEN aStation[nStation] := pStation; END_IF
END_METHOD

// Nouveau déploiement : états des calibrations retrouvés par identifiant
METHOD OnDeploy
VAR
    i : INT;
END_VAR
Abort();
FOR i := 1 TO GVL_Const.CALIB_PER_STATION DO
    IF i <= _refMachine.nCalibCount AND aCalib[i].nId <> _refMachine.aCalib[i].nId THEN
        MEMSET(ADR(aCalib[i]), 0, SIZEOF(aCalib[i]));
        aCalib[i].nId := _refMachine.aCalib[i].nId;
    END_IF
    IF i <= _refMachine.nCalibCount THEN aCalib[i].nValidityDays := _refMachine.aCalib[i].nValidityDays; END_IF
END_FOR
END_METHOD

METHOD Start : E_RejectReason
VAR_INPUT
    nTable : USINT;
    nMover : USINT;
    pMover : POINTER TO ST_MoverCtx;
    sUser : STRING(24);
END_VAR
VAR
    i : INT;
END_VAR
IF bRunning THEN Start := E_RejectReason.Busy; RETURN; END_IF
IF nTable < 1 OR nTable > GVL_Const.MAX_TABLES OR_ELSE NOT _refMachine.aTable[nTable].bUsed
   OR_ELSE _refMachine.aTable[nTable].eKind <> E_TableKind.MachineCalibration THEN
    Start := E_RejectReason.NotConfigured;
    RETURN;
END_IF
_nTable := nTable;
_nPC := _refMachine.aTable[nTable].nStart;
_nCalib := 0;
FOR i := 1 TO MIN(_refMachine.nCalibCount, GVL_Const.CALIB_PER_STATION) DO
    IF _refMachine.aCalib[i].nTable = nTable THEN _nCalib := INT_TO_USINT(i); END_IF
END_FOR
_nMover := nMover;
_pMover := pMover;
_sUser := sUser;
_nWait := 0;
_nRetry := 0;
_bAnswered := FALSE;
stPrompt.nPromptId := 0;
IF _nCalib > 0 THEN aCalib[_nCalib].eState := E_CalibState.Running; END_IF
bRunning := TRUE;
Start := E_RejectReason.None;
END_METHOD

METHOD Abort
IF bRunning THEN _Fail(0); END_IF
END_METHOD

METHOD AnswerPrompt : BOOL
VAR_INPUT
    nPromptId : UDINT;
    bConfirm : BOOL;
END_VAR
AnswerPrompt := FALSE;
IF stPrompt.nPromptId = 0 OR stPrompt.nPromptId <> nPromptId THEN RETURN; END_IF
_bAnswered := TRUE;
_bConfirm := bConfirm;
AnswerPrompt := TRUE;
END_METHOD

METHOD Cycle
VAR_INPUT
    bHmiLost : BOOL;
END_VAR
VAR
    nGuard : INT;
    ins : REFERENCE TO ST_Instr;
    st : POINTER TO FB_Station;
    nCalibTable : USINT;
    k : INT;
    eSev : E_Severity;
    aZero : ARRAY[1..GVL_Const.MAX_PARAMS] OF LREAL;
END_VAR
IF NOT bRunning THEN RETURN; END_IF
FOR nGuard := 1 TO GVL_Const.MAX_INSTR_PER_CYCLE DO
    IF _nPC < _refMachine.aTable[_nTable].nStart OR _nPC >= _refMachine.aTable[_nTable].nStart + _refMachine.aTable[_nTable].nLength THEN
        _Fail(905);
        RETURN;
    END_IF
    ins REF= _refMachine.aInstr[_nPC];
    CASE ins.eOp OF
        E_Op.Nop, E_Op.StepBegin, E_Op.StepEnd:
            _nPC := _nPC + 1;
        E_Op.Jump:
            _nPC := DINT_TO_INT(ins.aArg[1]);
        E_Op.WaitTime:
            IF _nWait = 0 THEN
                _nWait := 1;
                _fWaitMs := ins.aParam[1].fValue;
                _fElapsedMs := 0;
            END_IF
            _fElapsedMs := _fElapsedMs + F_CycleMs();
            IF _fElapsedMs < _fWaitMs THEN RETURN; END_IF
            _nWait := 0;
            _nPC := _nPC + 1;
        E_Op.Prompt:
            IF _nWait = 0 THEN
                _nWait := 3;
                _nPromptSeq := _nPromptSeq + 1;
                stPrompt.nPromptId := _nPromptSeq;
                stPrompt.nText := DINT_TO_INT(ins.aArg[1]);
                stPrompt.bInput := ins.aArg[2] = 1;
                _bAnswered := FALSE;
            END_IF
            IF bHmiLost OR (_bAnswered AND NOT _bConfirm) THEN
                stPrompt.nPromptId := 0;
                _nWait := 0;
                IF NOT _Failure(ins, 908) THEN RETURN; END_IF
            ELSIF _bAnswered THEN
                stPrompt.nPromptId := 0;
                _nWait := 0;
                _nPC := _nPC + 1;
            ELSE
                RETURN;
            END_IF
        E_Op.CalibStation:
            _nStation := DINT_TO_USINT(ins.aArg[1]);
            IF _nStation < 1 OR _nStation > GVL_Const.MAX_STATIONS OR_ELSE aStation[_nStation] = 0 THEN _Fail(905); RETURN; END_IF
            st := aStation[_nStation];
            IF _nWait = 0 THEN
                k := DINT_TO_INT(ins.aArg[2]);
                nCalibTable := 0;
                IF k >= 1 AND k <= GVL_Const.CALIB_PER_STATION THEN nCalibTable := st^.Data.aCalib[k].nTable; END_IF
                IF st^.Launch(nCalibTable, 0, 0, 0, aZero, _sUser) <> E_RejectReason.None THEN
                    IF NOT _Failure(ins, 909) THEN RETURN; END_IF
                ELSE
                    _nWait := 2;
                    RETURN;
                END_IF
            ELSIF st^.Response.eStatus = E_OpStatus.Done THEN
                st^.AckResponse();
                _nWait := 0;
                _nRetry := 0;
                _nPC := _nPC + 1;
            ELSIF st^.Response.eStatus = E_OpStatus.Failed OR st^.Response.eStatus = E_OpStatus.Aborted THEN
                st^.AckResponse();
                _nWait := 0;
                IF NOT _Failure(ins, 909) THEN RETURN; END_IF
            ELSE
                RETURN;
            END_IF
        E_Op.Route:
            IF NOT _Route(ins) THEN RETURN; END_IF
        E_Op.Alarm:
            IF ins.aArg[2] = 1 THEN eSev := E_Severity.Warning; ELSE eSev := E_Severity.MachineFault; END_IF
            IF __ISVALIDREF(_refAlarms) THEN _refAlarms.RaiseEvent(0, DINT_TO_UINT(ins.aArg[3]), DINT_TO_UDINT(ins.aArg[1]), eSev); END_IF
            IF ins.aArg[2] >= 2 THEN _Fail(0); RETURN; END_IF
            _nPC := _nPC + 1;
        E_Op.End:
            _Succeed();
            RETURN;
    ELSE
        _Fail(905);
        RETURN;
    END_CASE
END_FOR
END_METHOD

// Route du mover choisi : déplacement en position de travail d'une station de la fonction, puis lancement de
// l'opération sur la station (comme un lancement HMI) ; TRUE quand l'instruction est terminée
METHOD PRIVATE _Route : BOOL
VAR_INPUT
    ins : REFERENCE TO ST_Instr;
END_VAR
VAR
    g : DINT;
    s : USINT;
    k : INT;
    nTable : USINT;
    aParam : ARRAY[1..GVL_Const.MAX_PARAMS] OF LREAL;
    st : POINTER TO FB_Station;
END_VAR
_Route := FALSE;
IF _nMover = 0 OR _pMover = 0 THEN _Fail(905); RETURN; END_IF
g := ins.aArg[1];
IF _nWait = 0 THEN
    _nStation := 0;
    FOR s := 1 TO GVL_Const.MAX_STATIONS DO
        IF _nStation = 0 AND g >= 1 AND g <= GVL_Const.MAX_GROUPS AND_THEN (SHR(_refMachine.aGroup[g].nStationMask, s - 1) AND 1) = 1 THEN
            _nStation := s;
        END_IF
    END_FOR
    IF _nStation = 0 OR_ELSE aStation[_nStation] = 0 THEN _Fail(905); RETURN; END_IF
    _nDest := _refMachine.aStation[_nStation].nWorkPos;
    IF NOT _refMgr.MoveTo(_nMover, _nDest) THEN RETURN; END_IF      // position occupée : on réessaie
    _nWait := 4;
    RETURN;
END_IF
st := aStation[_nStation];
IF _nWait = 4 THEN
    IF _refMgr.Moving(_nMover) THEN RETURN; END_IF
    nTable := 0;
    FOR k := 1 TO st^.Data.nOpMapCount DO
        IF st^.Data.aOpMap[k].nGroup = DINT_TO_USINT(g) AND st^.Data.aOpMap[k].nOperationNo = DINT_TO_USINT(ins.aArg[2]) THEN nTable := st^.Data.aOpMap[k].nTable; END_IF
    END_FOR
    FOR k := 1 TO GVL_Const.MAX_PARAMS DO aParam[k] := ins.aParam[k].fValue; END_FOR
    IF st^.Launch(nTable, _nMover, _pMover, DINT_TO_USINT(ins.aArg[3]), aParam, _sUser) <> E_RejectReason.None THEN
        _nWait := 0;
        _Route := _Failure(ins, 909);
        RETURN;
    END_IF
    _nWait := 2;
    RETURN;
END_IF
IF st^.Response.eStatus = E_OpStatus.Done THEN
    st^.AckResponse();
    _nWait := 0;
    _nPC := _nPC + 1;
    _Route := TRUE;
ELSIF st^.Response.eStatus = E_OpStatus.Failed OR st^.Response.eStatus = E_OpStatus.Aborted THEN
    st^.AckResponse();
    _nWait := 0;
    _Route := _Failure(ins, 909);
END_IF
END_METHOD

// Politique d'échec de la carte (docs/05 § 3.6) ; TRUE si l'exécution continue ce cycle
METHOD PRIVATE _Failure : BOOL
VAR_INPUT
    ins : REFERENCE TO ST_Instr;
    nCode : UINT;
END_VAR
_Failure := FALSE;
CASE ins.eOnFail OF
    E_FailPolicy.Retry:
        IF _nRetry < ins.nRetries THEN
            _nRetry := _nRetry + 1;
            RETURN;                                     // même PC : relance au cycle suivant
        END_IF
        _Fail(nCode);
    E_FailPolicy.Ignore:
        _nRetry := 0;
        _nPC := _nPC + 1;
        _Failure := TRUE;
    E_FailPolicy.Goto:
        _nRetry := 0;
        _nPC := ins.nFailTarget;
        _Failure := TRUE;
ELSE
    _Fail(nCode);
END_CASE
END_METHOD

METHOD PRIVATE _Succeed
IF _nCalib > 0 THEN
    aCalib[_nCalib].eState := E_CalibState.Valid;
    aCalib[_nCalib].tLast := F_NowUtc();
    aCalib[_nCalib].sUser := _sUser;
END_IF
stPrompt.nPromptId := 0;
bRunning := FALSE;
END_METHOD

METHOD PRIVATE _Fail
VAR_INPUT
    nCode : UINT;
END_VAR
IF _nCalib > 0 THEN aCalib[_nCalib].eState := E_CalibState.Failed; END_IF
IF nCode <> 0 AND __ISVALIDREF(_refAlarms) THEN _refAlarms.RaiseEvent(0, nCode, INT_TO_UDINT(_nTable), E_Severity.Warning); END_IF
stPrompt.nPromptId := 0;
_nWait := 0;
bRunning := FALSE;
END_METHOD

// Calibrations machine échues ou jamais faites : avertissement 912 (docs/05 § 10.1)
METHOD CheckCalibrations
VAR_INPUT
    tNow : LINT;
END_VAR
VAR
    i : INT;
END_VAR
FOR i := 1 TO MIN(_refMachine.nCalibCount, GVL_Const.CALIB_PER_STATION) DO
    IF aCalib[i].eState = E_CalibState.Valid AND aCalib[i].nValidityDays > 0
       AND tNow - aCalib[i].tLast > UINT_TO_LINT(aCalib[i].nValidityDays) * 864000000000 THEN
        aCalib[i].eState := E_CalibState.Expired;
    END_IF
    IF (aCalib[i].eState = E_CalibState.Expired OR aCalib[i].eState = E_CalibState.Never) AND __ISVALIDREF(_refAlarms) THEN
        _refAlarms.RaiseEvent(0, 912, INT_TO_UDINT(i), E_Severity.Warning);
    END_IF
END_FOR
END_METHOD

METHOD PublishRetained
VAR_IN_OUT
    stOut : ST_RetainedValues;
END_VAR
VAR
    i : INT;
    stItem : ST_RetainedItem;
END_VAR
FOR i := 1 TO MIN(_refMachine.nCalibCount, GVL_Const.CALIB_PER_STATION) DO
    MEMSET(ADR(stItem), 0, SIZEOF(stItem));
    stItem.eKind := E_RetainedKind.Calibration;
    stItem.nId := aCalib[i].nId;
    stItem.aValue[1] := F_CalibStateNum(aCalib[i].eState);
    stItem.tStamp := aCalib[i].tLast;
    stItem.sUser := aCalib[i].sUser;
    F_AddRetained(stOut, stItem);
END_FOR
END_METHOD

METHOD Restore : BOOL
VAR_IN_OUT
    stItem : ST_RetainedItem;
END_VAR
VAR
    i : INT;
END_VAR
Restore := FALSE;
IF stItem.eKind <> E_RetainedKind.Calibration OR stItem.nId = 0 THEN RETURN; END_IF
FOR i := 1 TO MIN(_refMachine.nCalibCount, GVL_Const.CALIB_PER_STATION) DO
    IF aCalib[i].nId = stItem.nId THEN
        aCalib[i].eState := F_CalibStateOf(stItem.aValue[1]);
        aCalib[i].tLast := stItem.tStamp;
        aCalib[i].sUser := stItem.sUser;
        Restore := TRUE;
        RETURN;
    END_IF
END_FOR
END_METHOD

METHOD Publish
VAR_IN_OUT
    stStatus : ST_MachineStatus;
END_VAR
stStatus.nCalib := _refMachine.nCalibCount;
stStatus.aCalib := aCalib;
stStatus.stPrompt := stPrompt;
END_METHOD
END_FUNCTION_BLOCK

(* ---- FB_ManualChannel.st ---- *)
// Canal manuel d'une station ou de la machine (canal 0) (docs/05 § 7) : action, jog avec garde, acquittement,
// apprentissage. Conditions : mode Maintenance et hôte Stopped ; les droits sont contrôlés par la HMI.
FUNCTION_BLOCK FB_ManualChannel
VAR
    _nStation : USINT;              // 0 = machine
    _ipHost : I_ManualHost;
    _nLastSeq : UDINT;
    _nObject : UINT;                // objet de l'action en cours, 0 = aucune
    _bJog : BOOL;
    _nLastAlive : UDINT;
    _fQuietMs : LREAL;
    _eStateAtStart : E_State;
END_VAR

METHOD Init
VAR_INPUT
    nStation : USINT;
    ipHost : I_ManualHost;
END_VAR
_nStation := nStation;
_ipHost := ipHost;
END_METHOD

METHOD Cycle
VAR
    req : REFERENCE TO ST_ManualRequest;
    resp : REFERENCE TO ST_ManualResponse;
    ipObj : I_Object;
END_VAR
IF _ipHost = 0 OR _nStation > GVL_Const.MAX_STATIONS THEN RETURN; END_IF
req REF= GVL_Hmi.aManual[_nStation];
resp REF= GVL_Hmi.aManualResp[_nStation];

// Suivi de l'action en cours
IF _nObject <> 0 THEN
    ipObj := _ipHost.ObjectAt(_nObject);
    IF ipObj <> 0 THEN
        resp.eActStatus := ipObj.ActStatus;
        resp.nErrorCode := ipObj.Status.nErrorCode;
        resp.nSubCode := ipObj.Status.nSubCode;
        resp.stResults := ipObj.Results;
        IF _bJog THEN
            // Garde du jog : la HMI incrémente nJogAlive toutes les 100 ms bouton tenu
            IF GVL_Hmi.nJogAlive <> _nLastAlive THEN
                _nLastAlive := GVL_Hmi.nJogAlive;
                _fQuietMs := 0;
            ELSE
                _fQuietMs := _fQuietMs + F_CycleMs();
            END_IF
            IF _fQuietMs >= GVL_Const.JOG_GUARD_MS OR _ipHost.State <> _eStateAtStart THEN
                ipObj.Abort();
                _bJog := FALSE;
                _nObject := 0;
            END_IF
        ELSIF ipObj.ActStatus <> E_ActStatus.Busy THEN
            _nObject := 0;
        END_IF
    ELSE
        _nObject := 0;
    END_IF
END_IF

IF req.nSeq = _nLastSeq THEN RETURN; END_IF
_nLastSeq := req.nSeq;
resp.nSeq := req.nSeq;
resp.eReason := E_RejectReason.None;
resp.eResult := E_CmdResult.Rejected;
IF _ipHost.Mode <> E_Mode.Maintenance THEN resp.eReason := E_RejectReason.WrongMode; RETURN; END_IF
IF _ipHost.State <> E_State.Stopped THEN resp.eReason := E_RejectReason.WrongState; RETURN; END_IF
IF req.eKind <> E_ManualKind.TeachPosition AND (req.nObject < 1 OR req.nObject > GVL_Const.MAX_OBJ_PER_STATION) THEN
    resp.eReason := E_RejectReason.NotConfigured;
    RETURN;
END_IF
IF req.eKind <> E_ManualKind.TeachPosition THEN
    ipObj := _ipHost.ObjectAt(req.nObject);
    IF ipObj = 0 THEN resp.eReason := E_RejectReason.NotConfigured; RETURN; END_IF
END_IF

CASE req.eKind OF
    E_ManualKind.Action, E_ManualKind.JogStart:
        IF _nObject <> 0 THEN resp.eReason := E_RejectReason.Busy; RETURN; END_IF
        resp.eStart := ipObj.Start(req.nAction, req.stParams, TRUE);
        IF resp.eStart = E_StartResult.Accepted THEN
            _nObject := req.nObject;
            _bJog := req.eKind = E_ManualKind.JogStart;
            _nLastAlive := GVL_Hmi.nJogAlive;
            _fQuietMs := 0;
            _eStateAtStart := _ipHost.State;
            resp.eResult := E_CmdResult.Accepted;
        END_IF
        resp.eActStatus := ipObj.ActStatus;
        resp.stResults := ipObj.Results;
    E_ManualKind.JogStop:
        ipObj.Abort();
        _bJog := FALSE;
        _nObject := 0;
        resp.eResult := E_CmdResult.Accepted;
    E_ManualKind.Ack:
        ipObj.Ack();
        resp.eResult := E_CmdResult.Accepted;
    E_ManualKind.TeachPosition:
        resp.eResult := SEL(_Teach(req := req, stTaught => resp.stTaught), E_CmdResult.Rejected, E_CmdResult.Accepted);
        IF resp.eResult = E_CmdResult.Rejected THEN resp.eReason := E_RejectReason.NotConfigured; END_IF
END_CASE
END_METHOD

// Apprentissage : position actuelle des axes indiqués, composantes choisies (docs/05 § 7)
METHOD PRIVATE _Teach : BOOL
VAR_INPUT
    req : REFERENCE TO ST_ManualRequest;
END_VAR
VAR_OUTPUT
    stTaught : ST_Position;
END_VAR
VAR
    k : USINT;
    n : UINT;
    fValue : LREAL;
    pPos : POINTER TO ST_NamedPos;
    ipObj : I_Object;
END_VAR
_Teach := FALSE;
pPos := _ipHost.NamedPos(req.nTeachPos);
IF pPos = 0 THEN RETURN; END_IF
stTaught := pPos^.stPos;
FOR k := 1 TO 4 DO
    n := req.aTeachFrom[k];
    IF (SHR(req.nTeachMask, k - 1) AND 1) = 1 THEN
        ipObj := _ipHost.ObjectAt(n);
        IF ipObj <> 0 THEN
            fValue := ipObj.Status.aValue[1];
            CASE k OF
                1: stTaught.fX := fValue;
                2: stTaught.fY := fValue;
                3: stTaught.fZ := fValue;
                4: stTaught.fC := fValue;
            END_CASE
        END_IF
    END_IF
END_FOR
pPos^.stPos := stTaught;
pPos^.bTaught := TRUE;
_Teach := TRUE;
END_METHOD
END_FUNCTION_BLOCK

(* ---- FB_MoverManager.st ---- *)
// Gestionnaire de movers (docs/05 § 6) : occupation et réservation des positions planaires, envoi des
// déplacements au pilote planaire, détection des arrivées (fenêtre de position et à l'arrêt 50 ms), timeout.
FUNCTION_BLOCK FB_MoverManager IMPLEMENTS I_MoverMotion
VAR
    _refMachine : REFERENCE TO ST_MachineData;
    ipDriver : I_PlanarDriver;
    aOwner : ARRAY[1..GVL_Const.MAX_PLANAR_POS] OF USINT;         // mover propriétaire, 0 = libre
    _aDest : ARRAY[1..GVL_Const.MAX_MOVERS] OF INT;
    _aMoveMs : ARRAY[1..GVL_Const.MAX_MOVERS] OF LREAL;
    _aStillMs : ARRAY[1..GVL_Const.MAX_MOVERS] OF LREAL;
    _aTimeoutMs : ARRAY[1..GVL_Const.MAX_MOVERS] OF LREAL;
    _aArrived : ARRAY[1..GVL_Const.MAX_MOVERS] OF INT;           // position atteinte ce cycle, 0 sinon
    _aTimedOut : ARRAY[1..GVL_Const.MAX_MOVERS] OF BOOL;
    _fVelocity : LREAL := 1000.0;
    _fAcceleration : LREAL := 5000.0;
    _fWindow : LREAL := 0.1;
END_VAR

METHOD Init
VAR_INPUT
    refMachine : REFERENCE TO ST_MachineData;
    ipPlanar : I_PlanarDriver;
END_VAR
_refMachine REF= refMachine;
ipDriver := ipPlanar;
END_METHOD

// Paramètres du système planaire (type 13 : P1 vitesse, P2 accélération, P3 fenêtre)
METHOD Configure
VAR
    i : UINT;
END_VAR
FOR i := 1 TO _refMachine.nMachineObj DO
    IF _refMachine.aMachineObj[i].nType = GVL_Catalog.Type_PlanarSystem THEN
        IF _refMachine.aMachineObj[i].aParam[1] > 0 THEN _fVelocity := _refMachine.aMachineObj[i].aParam[1]; END_IF
        IF _refMachine.aMachineObj[i].aParam[2] > 0 THEN _fAcceleration := _refMachine.aMachineObj[i].aParam[2]; END_IF
        IF _refMachine.aMachineObj[i].aParam[3] > 0 THEN _fWindow := _refMachine.aMachineObj[i].aParam[3]; END_IF
    END_IF
END_FOR
END_METHOD

METHOD Owner : USINT
VAR_INPUT
    nPos : INT;
END_VAR
IF nPos >= 1 AND nPos <= GVL_Const.MAX_PLANAR_POS THEN Owner := aOwner[nPos]; END_IF
END_METHOD

METHOD Reserve
VAR_INPUT
    nPos : INT;
    nMover : USINT;
END_VAR
IF nPos >= 1 AND nPos <= GVL_Const.MAX_PLANAR_POS THEN aOwner[nPos] := nMover; END_IF
END_METHOD

METHOD Free
VAR_INPUT
    nPos : INT;
    nMover : USINT;
END_VAR
IF nPos >= 1 AND nPos <= GVL_Const.MAX_PLANAR_POS AND_THEN aOwner[nPos] = nMover THEN aOwner[nPos] := 0; END_IF
END_METHOD

// Libère toutes les positions d'un mover sauf nKeep
METHOD FreeAll
VAR_INPUT
    nMover : USINT;
    nKeep : INT;
END_VAR
VAR
    i : INT;
END_VAR
FOR i := 1 TO GVL_Const.MAX_PLANAR_POS DO
    IF aOwner[i] = nMover AND i <> nKeep THEN aOwner[i] := 0; END_IF
END_FOR
END_METHOD

// Réserve la destination puis envoie le déplacement (docs/05 § 6.2)
METHOD MoveTo : BOOL
VAR_INPUT
    nMover : USINT;
    nPos : INT;
END_VAR
VAR
    stCur : ST_Position;
    fDist : LREAL;
END_VAR
MoveTo := FALSE;
IF ipDriver = 0 OR nPos < 1 OR nPos > _refMachine.nPlanarPos OR nMover < 1 OR nMover > GVL_Const.MAX_MOVERS THEN RETURN; END_IF
IF aOwner[nPos] <> 0 AND aOwner[nPos] <> nMover THEN RETURN; END_IF
IF NOT ipDriver.MoveTo(nMover, _refMachine.aPlanarPos[nPos].stPos, _fVelocity, _fAcceleration) THEN RETURN; END_IF
FreeAll(nMover, 0);
aOwner[nPos] := nMover;
_aDest[nMover] := nPos;
_aMoveMs[nMover] := 0;
_aStillMs[nMover] := 0;
_aArrived[nMover] := 0;
_aTimedOut[nMover] := FALSE;
stCur := ipDriver.MoverPosition(nMover);
fDist := SQRT(EXPT(_refMachine.aPlanarPos[nPos].stPos.fX - stCur.fX, 2) + EXPT(_refMachine.aPlanarPos[nPos].stPos.fY - stCur.fY, 2));
_aTimeoutMs[nMover] := 2.0 * (fDist / _fVelocity + _fVelocity / _fAcceleration) * 1000.0 + 5000.0;
MoveTo := TRUE;
END_METHOD

METHOD Cycle
VAR_INPUT
    fOverride : LREAL;
END_VAR
VAR
    i : USINT;
    stPos : ST_Position;
    nPos : INT;
    fDt : LREAL;
END_VAR
IF ipDriver = 0 THEN RETURN; END_IF
ipDriver.Cycle(fOverride);
fDt := F_CycleMs();
FOR i := 1 TO _refMachine.nMovers DO
    _aArrived[i] := 0;
    nPos := _aDest[i];
    IF nPos > 0 THEN
        stPos := ipDriver.MoverPosition(i);
        IF fOverride > 0 THEN _aMoveMs[i] := _aMoveMs[i] + fDt * fOverride / 100.0; END_IF
        IF NOT ipDriver.MoverMoving(i)
           AND ABS(stPos.fX - _refMachine.aPlanarPos[nPos].stPos.fX) <= MAX(_fWindow, 0.01)
           AND ABS(stPos.fY - _refMachine.aPlanarPos[nPos].stPos.fY) <= MAX(_fWindow, 0.01) THEN
            _aStillMs[i] := _aStillMs[i] + fDt;
            IF _aStillMs[i] >= GVL_Const.ARRIVAL_SETTLE_MS THEN
                _aArrived[i] := nPos;
                _aDest[i] := 0;
            END_IF
        ELSE
            _aStillMs[i] := 0;
            IF _aMoveMs[i] > _aTimeoutMs[i] THEN
                _aTimedOut[i] := TRUE;
                _aDest[i] := 0;
            END_IF
        END_IF
    END_IF
END_FOR
END_METHOD

// Position atteinte ce cycle (0 sinon)
METHOD Arrived : INT
VAR_INPUT
    nMover : USINT;
END_VAR
IF nMover >= 1 AND nMover <= GVL_Const.MAX_MOVERS THEN Arrived := _aArrived[nMover]; END_IF
END_METHOD

METHOD TimedOut : BOOL
VAR_INPUT
    nMover : USINT;
END_VAR
TimedOut := nMover >= 1 AND nMover <= GVL_Const.MAX_MOVERS AND_THEN _aTimedOut[nMover];
END_METHOD

METHOD Moving : BOOL
VAR_INPUT
    nMover : USINT;
END_VAR
Moving := nMover >= 1 AND nMover <= GVL_Const.MAX_MOVERS AND_THEN (_aDest[nMover] <> 0 OR (ipDriver <> 0 AND_THEN ipDriver.MoverMoving(nMover)));
END_METHOD

// Mode manuel (docs/05 § 6.5) : le mover quitte ses positions ; arrivé sur une position planaire libre, il la tient
METHOD MoveFree : BOOL
VAR_INPUT
    nMover : USINT;
    stPos : ST_Position;
    fSpeedPct : LREAL;
END_VAR
VAR
    k : INT;
END_VAR
MoveFree := FALSE;
IF ipDriver = 0 OR nMover < 1 OR nMover > GVL_Const.MAX_MOVERS THEN RETURN; END_IF
// Une position planaire tenue par un autre mover ne peut pas être visée
FOR k := 1 TO _refMachine.nPlanarPos DO
    IF _Near(stPos, _refMachine.aPlanarPos[k].stPos) AND aOwner[k] <> 0 AND aOwner[k] <> nMover THEN RETURN; END_IF
END_FOR
IF NOT ipDriver.MoveTo(nMover, stPos, _fVelocity * LIMIT(1.0, fSpeedPct, 100.0) / 100.0, _fAcceleration) THEN RETURN; END_IF
FreeAll(nMover, 0);
_aDest[nMover] := 0;
_aTimedOut[nMover] := FALSE;
FOR k := 1 TO _refMachine.nPlanarPos DO
    IF _Near(stPos, _refMachine.aPlanarPos[k].stPos) THEN aOwner[k] := nMover; END_IF
END_FOR
MoveFree := TRUE;
END_METHOD

METHOD StopMover
VAR_INPUT
    nMover : USINT;
END_VAR
IF ipDriver <> 0 THEN ipDriver.StopMover(nMover); END_IF
IF nMover >= 1 AND nMover <= GVL_Const.MAX_MOVERS THEN _aDest[nMover] := 0; END_IF
END_METHOD

METHOD Position : ST_Position
VAR_INPUT
    nMover : USINT;
END_VAR
IF ipDriver <> 0 THEN Position := ipDriver.MoverPosition(nMover); END_IF
END_METHOD

METHOD PRIVATE _Near : BOOL
VAR_INPUT
    a : ST_Position;
    b : ST_Position;
END_VAR
_Near := ABS(a.fX - b.fX) <= MAX(_fWindow, 0.5) AND ABS(a.fY - b.fY) <= MAX(_fWindow, 0.5);
END_METHOD

METHOD AnyMoving : BOOL
VAR
    i : USINT;
END_VAR
AnyMoving := FALSE;
FOR i := 1 TO GVL_Const.MAX_MOVERS DO
    IF Moving(i) THEN AnyMoving := TRUE; END_IF
END_FOR
END_METHOD

// Arrêt contrôlé de tous les movers (Abort) : les destinations sont abandonnées, les réservations gardées
METHOD StopAll
VAR
    i : USINT;
END_VAR
IF ipDriver <> 0 THEN ipDriver.StopAll(); END_IF
FOR i := 1 TO GVL_Const.MAX_MOVERS DO _aDest[i] := 0; END_FOR
END_METHOD

// Position planaire connue où se trouve le mover (Reset machine, docs/05 § 6.3), 0 sinon
METHOD PositionAt : INT
VAR_INPUT
    nMover : USINT;
END_VAR
VAR
    i : INT;
    stPos : ST_Position;
END_VAR
PositionAt := 0;
IF ipDriver = 0 THEN RETURN; END_IF
stPos := ipDriver.MoverPosition(nMover);
FOR i := 1 TO _refMachine.nPlanarPos DO
    IF ABS(stPos.fX - _refMachine.aPlanarPos[i].stPos.fX) <= MAX(_fWindow, 0.5) AND ABS(stPos.fY - _refMachine.aPlanarPos[i].stPos.fY) <= MAX(_fWindow, 0.5) THEN
        PositionAt := i;
        RETURN;
    END_IF
END_FOR
END_METHOD

// Position tampon libre la plus proche du mover, 0 si aucune
METHOD NearestFree : INT
VAR_INPUT
    nMover : USINT;
    eKind : E_PlanarPosKind;
END_VAR
VAR
    i : INT;
    stPos : ST_Position;
    fD : LREAL;
    fBest : LREAL := 1.0E30;
END_VAR
NearestFree := 0;
IF ipDriver = 0 THEN RETURN; END_IF
stPos := ipDriver.MoverPosition(nMover);
FOR i := 1 TO _refMachine.nPlanarPos DO
    IF _refMachine.aPlanarPos[i].eKind = eKind AND (aOwner[i] = 0 OR aOwner[i] = nMover) THEN
        fD := ABS(_refMachine.aPlanarPos[i].stPos.fX - stPos.fX) + ABS(_refMachine.aPlanarPos[i].stPos.fY - stPos.fY);
        IF fD < fBest THEN
            fBest := fD;
            NearestFree := i;
        END_IF
    END_IF
END_FOR
END_METHOD

PROPERTY Driver : I_PlanarDriver
GET
Driver := ipDriver;
END_GET
END_PROPERTY
END_FUNCTION_BLOCK

(* ---- FB_PackML.st ---- *)
// Machine d'états PackML réduite, commune à la machine et aux stations (docs/05 § 2)
FUNCTION_BLOCK FB_PackML
VAR_INPUT
    eCmd : E_Cmd;                   // commande du cycle, None sinon
    bStateComplete : BOOL;          // le travail de l'état est fini
    bFault : BOOL;                  // défaut qui impose Aborted
END_VAR
VAR_OUTPUT
    eState : E_State := E_State.Stopped;
    bEntry : BOOL;                  // vrai au premier cycle dans un nouvel état
    eLastCmdResult : E_CmdResult;   // None si aucune commande ce cycle
    tSince : LINT;                  // heure d'entrée dans l'état (UTC)
END_VAR
VAR
    eNext : E_State;
END_VAR

bEntry := FALSE;
eNext := eState;
IF bFault AND eState <> E_State.Aborted THEN
    eNext := E_State.Aborted;
ELSE
    CASE eState OF
    E_State.Stopped:
        IF eCmd = E_Cmd.Reset THEN eNext := E_State.Resetting;
        ELSIF eCmd = E_Cmd.Abort THEN eNext := E_State.Aborted; END_IF
    E_State.Resetting:
        IF eCmd = E_Cmd.Abort THEN eNext := E_State.Aborted;
        ELSIF eCmd = E_Cmd.Stop THEN eNext := E_State.Stopping;
        ELSIF bStateComplete THEN eNext := E_State.Idle; END_IF
    E_State.Idle:
        IF eCmd = E_Cmd.Start THEN eNext := E_State.Execute;
        ELSIF eCmd = E_Cmd.Stop THEN eNext := E_State.Stopping;
        ELSIF eCmd = E_Cmd.Abort THEN eNext := E_State.Aborted; END_IF
    E_State.Execute:
        IF eCmd = E_Cmd.Hold THEN eNext := E_State.Held;
        ELSIF eCmd = E_Cmd.Stop THEN eNext := E_State.Stopping;
        ELSIF eCmd = E_Cmd.Abort THEN eNext := E_State.Aborted; END_IF
    E_State.Held:
        IF eCmd = E_Cmd.Start THEN eNext := E_State.Execute;
        ELSIF eCmd = E_Cmd.Stop THEN eNext := E_State.Stopping;
        ELSIF eCmd = E_Cmd.Abort THEN eNext := E_State.Aborted; END_IF
    E_State.Stopping:
        IF eCmd = E_Cmd.Abort THEN eNext := E_State.Aborted;
        ELSIF bStateComplete THEN eNext := E_State.Stopped; END_IF
    E_State.Aborted:
        IF eCmd = E_Cmd.Clear THEN eNext := E_State.Clearing; END_IF
    E_State.Clearing:
        IF eCmd = E_Cmd.Abort THEN eNext := E_State.Aborted;
        ELSIF bStateComplete THEN eNext := E_State.Stopped; END_IF
    END_CASE
END_IF
IF eCmd = E_Cmd.None OR eCmd = E_Cmd.DrainStart OR eCmd = E_Cmd.DrainCancel THEN
    eLastCmdResult := E_CmdResult.None;         // pas de commande PackML ce cycle
ELSE
    eLastCmdResult := SEL(eNext <> eState, E_CmdResult.Rejected, E_CmdResult.Accepted);
END_IF
IF eNext <> eState THEN
    eState := eNext;
    bEntry := TRUE;
    tSince := F_NowUtc();
END_IF

// Accepterait-on cette commande dans l'état courant ? (pour refuser avant de l'appliquer, sans changer d'état)
METHOD Accepts : BOOL
VAR_INPUT
    eCommand : E_Cmd;
END_VAR
CASE eCommand OF
    E_Cmd.Reset: Accepts := eState = E_State.Stopped;
    E_Cmd.Start: Accepts := eState = E_State.Idle OR eState = E_State.Held;
    E_Cmd.Hold: Accepts := eState = E_State.Execute;
    E_Cmd.Stop: Accepts := eState = E_State.Resetting OR eState = E_State.Idle OR eState = E_State.Execute OR eState = E_State.Held;
    E_Cmd.Abort: Accepts := eState <> E_State.Aborted;
    E_Cmd.Clear: Accepts := eState = E_State.Aborted;
ELSE
    Accepts := FALSE;
END_CASE
END_METHOD

// Remet l'automate à Stopped (déploiement, démarrage du PLC)
METHOD ForceStopped
eState := E_State.Stopped;
bEntry := TRUE;
tSince := F_NowUtc();
END_METHOD
END_FUNCTION_BLOCK

(* ---- FB_PlanarSim.st ---- *)
// Système planaire simulé (docs/06 § 8) : déplacement en ligne droite, profil en S, arrêt si la destination est occupée
// (l'occupation est gérée par FB_MoverManager, qui ne donne jamais une destination déjà prise).
FUNCTION_BLOCK FB_PlanarSim IMPLEMENTS I_PlanarDriver
VAR
    nMovers : USINT;
    _bActive : BOOL;
    _fActivateMs : LREAL;
    _aPos : ARRAY[1..GVL_Const.MAX_MOVERS] OF ST_Position;
    _aFrom : ARRAY[1..GVL_Const.MAX_MOVERS] OF ST_Position;
    _aTo : ARRAY[1..GVL_Const.MAX_MOVERS] OF ST_Position;
    _aT : ARRAY[1..GVL_Const.MAX_MOVERS] OF LREAL;          // 0..1 avancement
    _aDurMs : ARRAY[1..GVL_Const.MAX_MOVERS] OF LREAL;
    _aMoving : ARRAY[1..GVL_Const.MAX_MOVERS] OF BOOL;
    _aAbsent : ARRAY[1..GVL_Const.MAX_MOVERS] OF BOOL;      // essai : mover retiré du plan
    _nError : UINT;
END_VAR

METHOD Activate : BOOL
VAR_INPUT
    bEnable : BOOL;
END_VAR
IF NOT bEnable THEN
    _bActive := FALSE;
    _fActivateMs := 0;
ELSIF NOT _bActive THEN
    _fActivateMs := _fActivateMs + F_CycleMs();
    IF _fActivateMs >= 1500.0 THEN _bActive := TRUE; END_IF
END_IF
Activate := _bActive;
END_METHOD

METHOD MoveTo : BOOL
VAR_INPUT
    nMover : USINT;
    stPos : ST_Position;
    fVelocity : LREAL;
    fAcceleration : LREAL;
END_VAR
VAR
    fDist : LREAL;
    fV : LREAL;
    fA : LREAL;
    fAccDist : LREAL;
END_VAR
MoveTo := FALSE;
IF NOT _bActive OR nMover < 1 OR nMover > nMovers OR_ELSE _aAbsent[nMover] THEN RETURN; END_IF
_aFrom[nMover] := _aPos[nMover];
_aTo[nMover] := stPos;
fDist := SQRT((stPos.fX - _aPos[nMover].fX) * (stPos.fX - _aPos[nMover].fX) + (stPos.fY - _aPos[nMover].fY) * (stPos.fY - _aPos[nMover].fY));
fV := MAX(fVelocity, 1.0);
fA := MAX(fAcceleration, 1.0);
fAccDist := fV * fV / fA;
IF fDist >= fAccDist THEN
    _aDurMs[nMover] := ((fDist - fAccDist) / fV + 2.0 * fV / fA) * 1000.0;
ELSE
    _aDurMs[nMover] := 2.0 * SQRT(fDist / fA) * 1000.0;
END_IF
_aDurMs[nMover] := MAX(_aDurMs[nMover], 50.0);
_aT[nMover] := 0;
_aMoving[nMover] := TRUE;
MoveTo := TRUE;
END_METHOD

METHOD StopAll
VAR
    i : USINT;
END_VAR
FOR i := 1 TO GVL_Const.MAX_MOVERS DO _aMoving[i] := FALSE; END_FOR
END_METHOD

METHOD StopMover
VAR_INPUT
    nMover : USINT;
END_VAR
IF nMover >= 1 AND nMover <= GVL_Const.MAX_MOVERS THEN _aMoving[nMover] := FALSE; END_IF
END_METHOD

METHOD AckError
_nError := 0;
END_METHOD

METHOD Cycle
VAR_INPUT
    fOverride : LREAL;
END_VAR
VAR
    i : USINT;
    e : LREAL;
END_VAR
FOR i := 1 TO nMovers DO
    IF _aMoving[i] AND _bActive THEN
        _aT[i] := MIN(1.0, _aT[i] + F_CycleMs() * LIMIT(0.0, fOverride, 100.0) / 100.0 / _aDurMs[i]);
        e := _aT[i] * _aT[i] * (3.0 - 2.0 * _aT[i]);
        _aPos[i].fX := _aFrom[i].fX + (_aTo[i].fX - _aFrom[i].fX) * e;
        _aPos[i].fY := _aFrom[i].fY + (_aTo[i].fY - _aFrom[i].fY) * e;
        _aPos[i].fC := _aTo[i].fC;
        IF _aT[i] >= 1.0 THEN
            _aPos[i] := _aTo[i];
            _aMoving[i] := FALSE;
        END_IF
    END_IF
END_FOR
END_METHOD

METHOD MoverPosition : ST_Position
VAR_INPUT
    nMover : USINT;
END_VAR
IF nMover >= 1 AND nMover <= GVL_Const.MAX_MOVERS THEN MoverPosition := _aPos[nMover]; END_IF
END_METHOD

METHOD MoverMoving : BOOL
VAR_INPUT
    nMover : USINT;
END_VAR
MoverMoving := nMover >= 1 AND nMover <= GVL_Const.MAX_MOVERS AND_THEN _aMoving[nMover];
END_METHOD

METHOD MoverDetected : BOOL
VAR_INPUT
    nMover : USINT;
END_VAR
MoverDetected := _bActive AND nMover >= 1 AND nMover <= nMovers AND_THEN NOT _aAbsent[nMover];
END_METHOD

METHOD SetInitialPosition
VAR_INPUT
    nMover : USINT;
    stPos : ST_Position;
END_VAR
IF nMover >= 1 AND nMover <= GVL_Const.MAX_MOVERS THEN _aPos[nMover] := stPos; END_IF
END_METHOD

// Essai : retirer un mover du plan, ou provoquer une collision (docs/12 § 5)
METHOD SetAbsent
VAR_INPUT
    nMover : USINT;
    bAbsent : BOOL;
END_VAR
IF nMover >= 1 AND nMover <= GVL_Const.MAX_MOVERS THEN _aAbsent[nMover] := bAbsent; END_IF
END_METHOD

METHOD SetError
VAR_INPUT
    nCode : UINT;
END_VAR
_nError := nCode;
END_METHOD

// Nombre de movers posés sur le plan simulé (configuration machine)
METHOD SetMoverCount
VAR_INPUT
    nCount : USINT;
END_VAR
nMovers := MIN(nCount, GVL_Const.MAX_MOVERS);
END_METHOD

PROPERTY Active : BOOL
GET
Active := _bActive;
END_GET
END_PROPERTY

PROPERTY ErrorCode : UINT
GET
ErrorCode := _nError;
END_GET
END_PROPERTY

PROPERTY ErrorSubCode : UDINT
GET
ErrorSubCode := 0;
END_GET
END_PROPERTY
END_FUNCTION_BLOCK

(* ---- FB_QualityMonitor.st ---- *)
// Surveillance des rebuts (docs/10 § 9) : rebuts successifs et taux sur fenêtre glissante en nombre de résultats,
// par station (constatés et imputés), fonction, mover, machine, et budget de rebuts par OF.
// Les réactions sont rendues par les sorties ; le séquenceur général les applique.
FUNCTION_BLOCK FB_QualityMonitor
VAR_OUTPUT
    aStationHold : ARRAY[1..GVL_Const.MAX_STATIONS] OF BOOL;   // réaction « arrêt qualité de la station »
    aMoverOut : ARRAY[1..GVL_Const.MAX_MOVERS] OF BOOL;        // réaction « mover hors service »
    bLoadingLocked : BOOL;                                     // réaction « arrêt du chargement »
    bMachineStop : BOOL;                                       // impulsion : réaction « arrêter la machine »
    bAnyReaction : BOOL;                                       // balise bleu clignotant
END_VAR
VAR
    _refMachine : REFERENCE TO ST_MachineData;
    _refAlarms : REFERENCE TO FB_AlarmManager;
END_VAR
VAR PERSISTENT
    stTracks : ST_QualityStatus;
END_VAR

METHOD Init
VAR_INPUT
    refMachine : REFERENCE TO ST_MachineData;
    refAlarms : REFERENCE TO FB_AlarmManager;
END_VAR
_refMachine REF= refMachine;
_refAlarms REF= refAlarms;
END_METHOD

METHOD PRIVATE _Rule : ST_QualityRule
VAR_INPUT
    eScope : E_QualityScope;
    nIndex : INT;
END_VAR
_Rule := _refMachine.stQuality.aDefault[TO_INT(eScope)];
CASE eScope OF
    E_QualityScope.Station:
        IF nIndex >= 1 AND nIndex <= GVL_Const.MAX_STATIONS AND_THEN NOT _refMachine.stQuality.aStationInherits[nIndex] THEN
            _Rule := _refMachine.stQuality.aStationRule[nIndex];
        END_IF
    E_QualityScope.Group:
        IF nIndex >= 1 AND nIndex <= GVL_Const.MAX_GROUPS AND_THEN NOT _refMachine.stQuality.aGroupInherits[nIndex] THEN
            _Rule := _refMachine.stQuality.aGroupRule[nIndex];
        END_IF
END_CASE
END_METHOD

METHOD PRIVATE _Track : POINTER TO ST_QualityTrack
VAR_INPUT
    eScope : E_QualityScope;
    nIndex : INT;
END_VAR
CASE eScope OF
    E_QualityScope.Station: _Track := ADR(stTracks.aStation[LIMIT(1, nIndex, GVL_Const.MAX_STATIONS)]);
    E_QualityScope.StationImputed: _Track := ADR(stTracks.aStationImputed[LIMIT(1, nIndex, GVL_Const.MAX_STATIONS)]);
    E_QualityScope.Group: _Track := ADR(stTracks.aGroup[LIMIT(1, nIndex, GVL_Const.MAX_GROUPS)]);
    E_QualityScope.Mover: _Track := ADR(stTracks.aMover[LIMIT(1, nIndex, GVL_Const.MAX_MOVERS)]);
ELSE
    _Track := ADR(stTracks.stMachine);
END_CASE
END_METHOD

// Un résultat (docs/10 § 9, « À chaque résultat »)
METHOD Record
VAR_INPUT
    eScope : E_QualityScope;
    nIndex : INT;
    bBad : BOOL;
END_VAR
VAR
    t : REFERENCE TO ST_QualityTrack;
    r : ST_QualityRule;
    nOld : USINT;
    nConsecAct : USINT;
    fRate : LREAL;
    bActConsec : BOOL;
    bActRate : BOOL;
    bWarn : BOOL;
END_VAR
t REF= _Track(eScope, nIndex)^;
r := _Rule(eScope, nIndex);
IF r.nWindow = 0 THEN r.nWindow := 1; END_IF
// fenêtre glissante
IF t.nCount >= r.nWindow THEN
    nOld := INT_TO_USINT((USINT_TO_INT(t.nHead) + 256 - USINT_TO_INT(t.nCount)) MOD 256);
    IF _Bit(t, nOld) AND t.nBadInWindow > 0 THEN t.nBadInWindow := t.nBadInWindow - 1; END_IF
ELSE
    t.nCount := t.nCount + 1;
END_IF
_SetBit(t, t.nHead, bBad);
t.nHead := INT_TO_USINT((USINT_TO_INT(t.nHead) + 1) MOD 256);
IF bBad THEN
    t.nBadInWindow := t.nBadInWindow + 1;
    IF t.nConsec < 255 THEN t.nConsec := t.nConsec + 1; END_IF
    t.nTotalBad := t.nTotalBad + 1;
ELSE
    t.nConsec := 0;
    t.nTotalGood := t.nTotalGood + 1;
END_IF
// évaluation
nConsecAct := SEL(t.nProbationLeft > 0, r.nConsecAction, 2);
IF t.nCount >= r.nMinSample AND t.nCount > 0 THEN fRate := 100.0 * USINT_TO_LREAL(t.nBadInWindow) / USINT_TO_LREAL(t.nCount); ELSE fRate := -1.0; END_IF
bActConsec := nConsecAct > 0 AND t.nConsec >= nConsecAct;
bActRate := r.fRateAction > 0 AND fRate >= r.fRateAction AND t.nProbationLeft = 0;
bWarn := (r.nConsecWarn > 0 AND t.nConsec >= r.nConsecWarn) OR (r.fRateWarn > 0 AND fRate >= r.fRateWarn);
IF t.nProbationLeft > 0 THEN t.nProbationLeft := t.nProbationLeft - 1; END_IF

IF (bActConsec OR bActRate) AND NOT t.bLocked THEN
    t.bLocked := TRUE;
    t.eLevel := E_QualityLevel.Action;
    _React(eScope, nIndex, SEL(bActConsec, r.eReactionRate, r.eReactionConsec));
    _RaiseAlarm(eScope, nIndex, bActConsec, E_Severity.Quality, SEL(bActConsec, LREAL_TO_UDINT(MAX(fRate, 0.0) * 10.0), USINT_TO_UDINT(t.nConsec)));
ELSIF bWarn AND t.eLevel = E_QualityLevel.Normal THEN
    t.eLevel := E_QualityLevel.Warning;
    _RaiseAlarm(eScope, nIndex, t.nConsec >= r.nConsecWarn AND r.nConsecWarn > 0, E_Severity.Warning, USINT_TO_UDINT(t.nConsec));
ELSIF NOT bWarn AND t.eLevel = E_QualityLevel.Warning THEN
    t.eLevel := SEL(t.nProbationLeft > 0, E_QualityLevel.Normal, E_QualityLevel.Probation);
ELSIF t.eLevel = E_QualityLevel.Probation AND t.nProbationLeft = 0 AND NOT t.bLocked THEN
    t.eLevel := E_QualityLevel.Normal;
END_IF
END_METHOD

// Budget de rebuts de l'OF (docs/10 § 4.3) : avertissement à 80 %, arrêt du chargement à 100 %
METHOD RecordOrder
VAR_INPUT
    refOrder : REFERENCE TO ST_OrderState;
    bBad : BOOL;
END_VAR
VAR
    fBudget : LREAL;
    fUsed : LREAL;
END_VAR
IF bBad THEN refOrder.stQuality.nTotalBad := refOrder.stQuality.nTotalBad + 1; ELSE refOrder.stQuality.nTotalGood := refOrder.stQuality.nTotalGood + 1; END_IF
IF _refMachine.stQuality.nOrderBudgetCount > 0 THEN
    fBudget := UDINT_TO_LREAL(_refMachine.stQuality.nOrderBudgetCount);
ELSIF _refMachine.stQuality.fOrderBudgetPct > 0 THEN
    fBudget := UDINT_TO_LREAL(refOrder.nQuantity) * REAL_TO_LREAL(_refMachine.stQuality.fOrderBudgetPct) / 100.0;
ELSE
    RETURN;
END_IF
IF fBudget <= 0 THEN RETURN; END_IF
fUsed := 100.0 * UDINT_TO_LREAL(refOrder.stQuality.nTotalBad) / fBudget;
IF fUsed >= 100.0 AND NOT refOrder.stQuality.bLocked THEN
    refOrder.stQuality.bLocked := TRUE;
    refOrder.stQuality.eLevel := E_QualityLevel.Action;
    bLoadingLocked := TRUE;
    bAnyReaction := TRUE;
    IF __ISVALIDREF(_refAlarms) THEN _refAlarms.Raise(0, 958, LREAL_TO_UDINT(fUsed * 10.0), E_Severity.Quality); END_IF
ELSIF fUsed >= 80.0 AND refOrder.stQuality.eLevel = E_QualityLevel.Normal THEN
    refOrder.stQuality.eLevel := E_QualityLevel.Warning;
    IF __ISVALIDREF(_refAlarms) THEN _refAlarms.Raise(0, 958, LREAL_TO_UDINT(fUsed * 10.0), E_Severity.Warning); END_IF
END_IF
END_METHOD

// Libération (docs/10 § 6) : remise à zéro de la portée, surveillance renforcée pour 10 résultats
METHOD Release : BOOL
VAR_INPUT
    eScope : E_QualityScope;
    nIndex : INT;
END_VAR
VAR
    t : REFERENCE TO ST_QualityTrack;
END_VAR
t REF= _Track(eScope, nIndex)^;
Release := t.bLocked;
IF NOT t.bLocked THEN RETURN; END_IF
_Clear(t);
t.nProbationLeft := 10;
t.eLevel := E_QualityLevel.Probation;
t.bLocked := FALSE;
CASE eScope OF
    E_QualityScope.Station, E_QualityScope.StationImputed:
        IF nIndex >= 1 AND nIndex <= GVL_Const.MAX_STATIONS THEN aStationHold[nIndex] := stTracks.aStation[nIndex].bLocked OR stTracks.aStationImputed[nIndex].bLocked; END_IF
    E_QualityScope.Mover:
        IF nIndex >= 1 AND nIndex <= GVL_Const.MAX_MOVERS THEN aMoverOut[nIndex] := FALSE; END_IF
    E_QualityScope.Group, E_QualityScope.Machine:
        bLoadingLocked := FALSE;
END_CASE
IF __ISVALIDREF(_refAlarms) THEN _refAlarms.Clear(_AlarmSource(eScope, nIndex), _AlarmCode(eScope, nIndex, TRUE)); _refAlarms.Clear(_AlarmSource(eScope, nIndex), _AlarmCode(eScope, nIndex, FALSE)); END_IF
_UpdateAny();
END_METHOD

// Remise à zéro manuelle d'une portée (droit quality.reset)
METHOD Reset
VAR_INPUT
    eScope : E_QualityScope;
    nIndex : INT;
END_VAR
VAR
    t : REFERENCE TO ST_QualityTrack;
END_VAR
t REF= _Track(eScope, nIndex)^;
_Clear(t);
t.eLevel := E_QualityLevel.Normal;
END_METHOD

// Changement de référence produit (D87) : toutes les portées repartent de zéro, sauf les verrous en cours
METHOD ResetAllWindows
VAR
    i : INT;
END_VAR
FOR i := 1 TO GVL_Const.MAX_STATIONS DO _Clear(stTracks.aStation[i]); _Clear(stTracks.aStationImputed[i]); END_FOR
FOR i := 1 TO GVL_Const.MAX_GROUPS DO _Clear(stTracks.aGroup[i]); END_FOR
FOR i := 1 TO GVL_Const.MAX_MOVERS DO _Clear(stTracks.aMover[i]); END_FOR
_Clear(stTracks.stMachine);
END_METHOD

METHOD Publish
GVL_Hmi.stQuality := stTracks;
GVL_Hmi.stQuality.bLoadingLocked := bLoadingLocked;
bMachineStop := FALSE;
END_METHOD

METHOD PRIVATE _Clear
VAR_IN_OUT
    t : ST_QualityTrack;
END_VAR
t.nConsec := 0;
MEMSET(ADR(t.aWindow), 0, SIZEOF(t.aWindow));
t.nHead := 0;
t.nCount := 0;
t.nBadInWindow := 0;
END_METHOD

METHOD PRIVATE _React
VAR_INPUT
    eScope : E_QualityScope;
    nIndex : INT;
    eReaction : E_QualityReaction;
END_VAR
CASE eReaction OF
    E_QualityReaction.StationHold:
        IF (eScope = E_QualityScope.Station OR eScope = E_QualityScope.StationImputed) AND nIndex >= 1 AND nIndex <= GVL_Const.MAX_STATIONS THEN aStationHold[nIndex] := TRUE; END_IF
    E_QualityReaction.MoverOut:
        IF eScope = E_QualityScope.Mover AND nIndex >= 1 AND nIndex <= GVL_Const.MAX_MOVERS THEN aMoverOut[nIndex] := TRUE; END_IF
    E_QualityReaction.StopLoading:
        bLoadingLocked := TRUE;
    E_QualityReaction.MachineStop:
        bMachineStop := TRUE;
END_CASE
_UpdateAny();
END_METHOD

METHOD PRIVATE _UpdateAny
VAR
    i : INT;
END_VAR
bAnyReaction := bLoadingLocked;
FOR i := 1 TO GVL_Const.MAX_STATIONS DO bAnyReaction := bAnyReaction OR aStationHold[i]; END_FOR
FOR i := 1 TO GVL_Const.MAX_MOVERS DO bAnyReaction := bAnyReaction OR aMoverOut[i]; END_FOR
bAnyReaction := bAnyReaction OR stTracks.stMachine.bLocked;
END_METHOD

// Codes 950 à 958 (docs/10 § 8, docs/14 § 3.1)
METHOD PRIVATE _AlarmCode : UINT
VAR_INPUT
    eScope : E_QualityScope;
    nIndex : INT;
    bConsec : BOOL;
END_VAR
CASE eScope OF
    E_QualityScope.Station: _AlarmCode := SEL(bConsec, 951, 950);
    E_QualityScope.StationImputed: _AlarmCode := SEL(bConsec, 953, 952);
    E_QualityScope.Group: _AlarmCode := 954;
    E_QualityScope.Mover: _AlarmCode := 955;
    E_QualityScope.Machine: _AlarmCode := SEL(bConsec, 957, 956);
ELSE
    _AlarmCode := 958;
END_CASE
END_METHOD

METHOD PRIVATE _AlarmSource : UDINT
VAR_INPUT
    eScope : E_QualityScope;
    nIndex : INT;
END_VAR
// station : n° de station × 1000 ; fonction, mover : 0 (machine), le sous-code et le contexte précisent
IF (eScope = E_QualityScope.Station OR eScope = E_QualityScope.StationImputed) AND nIndex >= 1 THEN
    _AlarmSource := INT_TO_UDINT(nIndex) * 1000;
ELSE
    _AlarmSource := 0;
END_IF
END_METHOD

METHOD PRIVATE _RaiseAlarm
VAR_INPUT
    eScope : E_QualityScope;
    nIndex : INT;
    bConsec : BOOL;
    eSeverity : E_Severity;
    nValue : UDINT;
END_VAR
VAR
    stCtx : ST_AlarmContext;
END_VAR
IF NOT __ISVALIDREF(_refAlarms) THEN RETURN; END_IF
IF eScope = E_QualityScope.Mover THEN stCtx.nMover := INT_TO_USINT(nIndex); _refAlarms.SetContext(stCtx); END_IF
_refAlarms.Raise(_AlarmSource(eScope, nIndex), _AlarmCode(eScope, nIndex, bConsec), nValue, eSeverity);
END_METHOD

METHOD PRIVATE _Bit : BOOL
VAR_IN_OUT
    t : ST_QualityTrack;
END_VAR
VAR_INPUT
    n : USINT;
END_VAR
_Bit := (SHR(t.aWindow[n / 8], n MOD 8) AND 1) = 1;
END_METHOD

METHOD PRIVATE _SetBit
VAR_IN_OUT
    t : ST_QualityTrack;
END_VAR
VAR_INPUT
    n : USINT;
    b : BOOL;
END_VAR
IF b THEN
    t.aWindow[n / 8] := t.aWindow[n / 8] OR SHL(BYTE#1, n MOD 8);
ELSE
    t.aWindow[n / 8] := t.aWindow[n / 8] AND NOT SHL(BYTE#1, n MOD 8);
END_IF
END_METHOD
END_FUNCTION_BLOCK
